(* IEC 61131-3 sources: Industry-PLC-LLM/data/PLCBEAD_repo/PLCBEAD_PLCEmbed-main/PLC-BEAD/Source/PLC_Programs (part 14) *)

(* ---- V3_XPRO.ST ---- *)
TYPE oscat_vector_3 :
	STRUCT
		X : REAL;
		Y : REAL;
		Z : REAL;
	END_STRUCT;
END_TYPE

FUNCTION_BLOCK V3_XPRO_Block
	VAR_INPUT
		A :	oscat_vector_3;
		B :	oscat_vector_3;
	END_VAR

	VAR_OUTPUT
		V3_XPRO :	oscat_vector_3;
	END_VAR

	V3_XPRO.X := A.Y * B.Z - A.Z * B.Y;
	V3_XPRO.Y := A.Z * B.X - A.X * B.Z;
	V3_XPRO.Z := A.X * B.Y - A.Y * B.X;

END_FUNCTION_BLOCK

PROGRAM program0
  	VAR
		A :	oscat_vector_3;
		B :	oscat_vector_3;
		V3_XPRO :	oscat_vector_3;
		func_block : V3_XPRO_Block;
  	END_VAR
	func_block.A := A;
	func_block.B := B;
	func_block();
	V3_XPRO := func_block.V3_XPRO;
END_PROGRAM

CONFIGURATION Config0
  RESOURCE Res0 ON PLC
    TASK task0(INTERVAL := T#20ms,PRIORITY := 0);
    PROGRAM instance0 WITH task0 : program0;
  END_RESOURCE
END_CONFIGURATION

(* ---- V3_YANG.ST ---- *)
TYPE oscat_vector_3:
  	STRUCT
		X : REAL;
		Y : REAL;
		Z : REAL;
  	END_STRUCT;
END_TYPE

FUNCTION_BLOCK V3_ABS_Block

	VAR_INPUT
		A :	oscat_vector_3;
	END_VAR

	VAR_OUTPUT
		V3_ABS :	REAL;
	END_VAR

	V3_ABS := SQRT(A.X * A.X + A.Y * A.Y + A.Z * A.Z);

END_FUNCTION_BLOCK

FUNCTION_BLOCK V3_YANG_Block
	VAR_INPUT
		A :	oscat_vector_3;
	END_VAR

	VAR_OUTPUT
		V3_YANG :	REAL;
	END_VAR

	VAR
		la :	REAL;
		V3_ABS :	V3_ABS_Block;
	END_VAR

	V3_ABS(A:=A);
	la:=V3_ABS.V3_ABS;

	IF la > 0.0 THEN
		V3_YANG := ACOS(A.Y / la);
	ELSE
		V3_YANG := 0.0;
	END_IF;

END_FUNCTION_BLOCK

PROGRAM program0
  	VAR
		A :	oscat_vector_3;
		V3_YANG :	REAL;
		func_block : V3_YANG_Block;
  	END_VAR
	func_block.A := A;
	func_block();
	V3_YANG := func_block.V3_YANG;
END_PROGRAM

CONFIGURATION Config0
  RESOURCE Res0 ON PLC
    TASK task0(INTERVAL := T#20ms,PRIORITY := 0);
    PROGRAM instance0 WITH task0 : program0;
  END_RESOURCE
END_CONFIGURATION

(* ---- V3_ZANG.ST ---- *)
TYPE oscat_vector_3:
  STRUCT
	X : REAL;
	Y : REAL;
	Z : REAL;
  END_STRUCT;
END_TYPE

FUNCTION_BLOCK V3_ABS_Block

	VAR_INPUT
		A :	oscat_vector_3;
	END_VAR

	VAR_OUTPUT
		V3_ABS :	REAL;
	END_VAR

	V3_ABS := SQRT(A.X * A.X + A.Y * A.Y + A.Z * A.Z);

END_FUNCTION_BLOCK

FUNCTION_BLOCK V3_ZANG_Block
	VAR_INPUT
		A :	oscat_vector_3;
	END_VAR

	VAR_OUTPUT
		V3_ZANG :	REAL;
	END_VAR

	VAR
		la :	REAL;
		V3_ABS :	V3_ABS_Block;
	END_VAR

	V3_ABS(A:=A);
	la:=V3_ABS.V3_ABS;

	IF la > 0.0 THEN
		V3_ZANG := ACOS(A.Z / la);
	ELSE
		V3_ZANG := 0.0;
	END_IF;

END_FUNCTION_BLOCK

PROGRAM program0
  	VAR
		A :	oscat_vector_3;
		V3_ZANG :	REAL;
		func_block : V3_ZANG_Block;
  	END_VAR
	func_block.A := A;
	func_block();
	V3_ZANG := func_block.V3_ZANG;
END_PROGRAM

CONFIGURATION Config0
  RESOURCE Res0 ON PLC
    TASK task0(INTERVAL := T#20ms,PRIORITY := 0);
    PROGRAM instance0 WITH task0 : program0;
  END_RESOURCE
END_CONFIGURATION

(* ---- WATER_CP.ST ---- *)
TYPE
	oscat_ARRAY_X               : ARRAY [0..1]    OF REAL;
	oscat_XY                    : ARRAY [1..20]   OF oscat_ARRAY_X := [0,0,0,0,0,0,0,0,0,0,0,0,0,0,0,0,0,0,0,0];
END_TYPE

FUNCTION_BLOCK LINEAR_INT_Block

	VAR_INPUT
		X :	REAL;
		XY :	oscat_XY;
		PTS :	INT;
	END_VAR

	VAR_OUTPUT
		LINEAR_INT :	REAL;
	END_VAR

	VAR
		i :	INT;
		i2 :	INT;
	END_VAR

	pts := MIN(pts,20);

	i := 2;

	WHILE (i < pts) AND (XY[i][0] < X) DO
		i := i + 1;
	END_WHILE;

	i2 := i-1;

	LINEAR_INT := ((XY[i][1] - XY[i2][1]) * X - XY[i][1] * XY[i2][0] + XY[i2][1] * XY[i][0]) / (XY[i][0] - XY[i2][0]);

END_FUNCTION_BLOCK

FUNCTION_BLOCK WATER_CP_Block

    VAR_INPUT
        T :	REAL;
    END_VAR

    VAR_OUTPUT
        CAP :	REAL;
    END_VAR

    VAR
        Pts :	INT;
        data :	oscat_XY;
        FB_LINEAR_INT :	LINEAR_INT_Block;
    END_VAR

    IF Pts = 0 THEN
        Pts := 10;

        data[01][0] := REAL#0.0;
        data[01][1] := REAL#4.228;
        data[02][0] := REAL#05.0;
        data[02][1] := REAL#4.200;
        data[03][0] := REAL#10.0;
        data[03][1] := REAL#4.188;
        data[04][0] := REAL#15.0;
        data[04][1] := REAL#4.184;
        data[05][0] := REAL#50.0;
        data[05][1] := REAL#4.181;
        data[06][0] := REAL#60.0;
        data[06][1] := REAL#4.183;
        data[07][0] := REAL#70.0;
        data[07][1] := REAL#4.187;
        data[08][0] := REAL#80.0;
        data[08][1] := REAL#4.194;
        data[09][0] := REAL#90.0;
        data[09][1] := REAL#4.204;
        data[10][0] := REAL#100.0;
        data[10][1] := REAL#4.220;

    END_IF;

    FB_LINEAR_INT(X:=T,XY:=Data,Pts:=Pts);
    cap:=FB_LINEAR_INT.LINEAR_INT;

END_FUNCTION_BLOCK

PROGRAM program0
	VAR
		T :	REAL;
        CAP :	REAL;

		func_block : WATER_CP_Block;
	END_VAR
	func_block.T := T;

	func_block();
	CAP  := func_block.CAP;
END_PROGRAM

CONFIGURATION Config0
	RESOURCE Res0 ON PLC
		TASK task0(INTERVAL := T#20ms,PRIORITY := 0);
		PROGRAM instance0 WITH task0 : program0;
	END_RESOURCE
END_CONFIGURATION

(* ---- WATER_ENTHALPY.ST ---- *)
TYPE
	oscat_ARRAY_X               : ARRAY [0..1]    OF REAL;
	oscat_XY                    : ARRAY [1..20]   OF oscat_ARRAY_X := [0,0,0,0,0,0,0,0,0,0,0,0,0,0,0,0,0,0,0,0];
END_TYPE

FUNCTION_BLOCK LINEAR_INT_Block

	VAR_INPUT
		X :	REAL;
		XY :	oscat_XY;
		PTS :	INT;
	END_VAR

	VAR_OUTPUT
		LINEAR_INT :	REAL;
	END_VAR

	VAR
		i :	INT;
		i2 :	INT;
	END_VAR

	pts := MIN(pts,20);

	i := 2;

	WHILE (i < pts) AND (XY[i][0] < X) DO
		i := i + 1;
	END_WHILE;

	i2 := i-1;

	LINEAR_INT := ((XY[i][1] - XY[i2][1]) * X - XY[i][1] * XY[i2][0] + XY[i2][1] * XY[i][0]) / (XY[i][0] - XY[i2][0]);

END_FUNCTION_BLOCK

FUNCTION_BLOCK WATER_ENTHALPY_Block

    VAR_INPUT
        T :	REAL;
    END_VAR

    VAR_OUTPUT
        RESULT :	REAL;
    END_VAR

    VAR
        Pts :	INT;
        data :	oscat_XY;
        FB_LINEAR_INT :	LINEAR_INT_Block;
    END_VAR

    IF Pts = 0 THEN
        Pts := 11;
        data[01][0] := REAL#0.0;
        data[01][1] := REAL#0.06;
        data[02][0] := REAL#10.0;
        data[02][1] := REAL#42.1;
        data[03][0] := REAL#20.0;
        data[03][1] := REAL#83.9;
        data[04][0] := REAL#30.0;
        data[04][1] := REAL#125.8;
        data[05][0] := REAL#40.0;
        data[05][1] := REAL#167.58;
        data[06][0] := REAL#50.0;
        data[06][1] := REAL#209.4;
        data[07][0] := REAL#60.0;
        data[07][1] := REAL#251.2;
        data[08][0] := REAL#70.0;
        data[08][1] := REAL#293.1;
        data[09][0] := REAL#80.0;
        data[09][1] := REAL#335.0;
        data[10][0] := REAL#90.0;
        data[10][1] := REAL#377.0;
        data[11][0] := REAL#100.0;
        data[11][1] := REAL#419.1;
    END_IF;

    FB_LINEAR_INT(X:=T,XY:=Data,Pts:=Pts);
    Result :=FB_LINEAR_INT.LINEAR_INT;

END_FUNCTION_BLOCK

PROGRAM program0
	VAR
		T :	REAL;
		RESULT :	REAL;

		func_block : WATER_ENTHALPY_Block;
	END_VAR
	func_block.T := T;

	func_block();
	RESULT  := func_block.RESULT;
END_PROGRAM

CONFIGURATION Config0
	RESOURCE Res0 ON PLC
		TASK task0(INTERVAL := T#20ms,PRIORITY := 0);
		PROGRAM instance0 WITH task0 : program0;
	END_RESOURCE
END_CONFIGURATION

(* ---- WEEKDAY_TO_STRING.ST ---- *)
TYPE
	oscat_STRING2 : STRING;
	oscat_STRING10 : STRING;
END_TYPE

TYPE oscat_HOLIDAY_DATA :
	STRUCT
		NAME : STRING;
		DAY : SINT;
		MONTH : SINT;
		USE : SINT;
		PAD_BYTE : BYTE;
	END_STRUCT;
END_TYPE

TYPE
	oscat_HOLIDAY_DATA_0_29 	: ARRAY [0..29] OF oscat_HOLIDAY_DATA;
END_TYPE

TYPE
	oscat_ELEMENT_WEEKDAYS	: ARRAY [1..7] OF oscat_STRING10;
  	oscat_WEEKDAYS			: ARRAY [1..3] OF oscat_ELEMENT_WEEKDAYS := [0,0,0];
	oscat_ELEMENT_WEEKDAYS2	: ARRAY [1..7] OF oscat_STRING2;
  	oscat_WEEKDAYS2			: ARRAY [1..3] OF oscat_ELEMENT_WEEKDAYS2 := [0,0,0];
END_TYPE

TYPE oscat_LANGUAGE:
  STRUCT
    DEFAULT 	: INT;
	LMAX    	: INT;
  END_STRUCT;
END_TYPE

FUNCTION_BLOCK SETUP_HOLIDAY_FR_Block

	VAR_IN_OUT
		HD :	oscat_HOLIDAY_DATA_0_29;
	END_VAR

	VAR
		init :	BOOL;
	END_VAR

	IF init THEN RETURN; END_IF;

	init := TRUE;

	HD[00].NAME := 'Nouve an';
	HD[00].DAY  := SINT#01;
	HD[00].MONTH := SINT#01;
	HD[00].USE := SINT#01;

	HD[01].NAME := 'St Valentin';
	HD[01].DAY  := SINT#14;
	HD[01].MONTH := SINT#02;
	HD[01].USE := SINT#00;

	HD[02].NAME := 'Vendredi Saint (alsace)';
	HD[02].DAY  := SINT#-2;
	HD[02].MONTH := SINT#00;
	HD[02].USE := SINT#00;

	HD[03].NAME := 'Dimanche de pques';
	HD[03].DAY  := SINT#00;
	HD[03].MONTH := SINT#00;
	HD[03].USE := SINT#01;

	HD[04].NAME := 'Lundi de pques';
	HD[04].DAY  := SINT#01;
	HD[04].MONTH := SINT#00;
	HD[04].USE := SINT#01;

	HD[05].NAME := 'Jeudi de Ascension';
	HD[05].DAY  := SINT#39;
	HD[05].MONTH := SINT#00;
	HD[05].USE := SINT#01;

	HD[06].NAME := 'dimanche de Pentecte';
	HD[06].DAY  := SINT#49;
	HD[06].MONTH := SINT#00;
	HD[06].USE := SINT#01;

	HD[07].NAME := 'jeudi de la Trinit';
	HD[07].DAY  := SINT#60;
	HD[07].MONTH := SINT#00;
	HD[07].USE := SINT#00;

	HD[08].NAME := 'Fte du travail';
	HD[08].DAY  := SINT#01;
	HD[08].MONTH := SINT#05;
	HD[08].USE := SINT#01;

	HD[09].NAME := 'Victoire 1945 ';
	HD[09].DAY  := SINT#08;
	HD[09].MONTH := SINT#05;
	HD[09].USE := SINT#01;

	HD[10].NAME := 'Prise de La bastille';
	HD[10].DAY  := SINT#14;
	HD[10].MONTH := SINT#07;
	HD[10].USE := SINT#01;

	HD[11].NAME := '15 Aot 1944';
	HD[11].DAY  := SINT#15;
	HD[11].MONTH := SINT#08;
	HD[11].USE := SINT#01;

	HD[12].NAME := 'Halloween';
	HD[12].DAY  := SINT#31;
	HD[12].MONTH := SINT#10;
	HD[12].USE := SINT#00;

	HD[13].NAME := 'Armistice 1918';
	HD[13].DAY  := SINT#11;
	HD[13].MONTH := SINT#11;
	HD[13].USE := SINT#01;

	HD[14].NAME := 'Nol';
	HD[14].DAY  := SINT#25;
	HD[14].MONTH := SINT#12;
	HD[14].USE := SINT#01;

	HD[15].NAME := 'Saint tienne (alsace)';
	HD[15].DAY  := SINT#26;
	HD[15].MONTH := SINT#12;
	HD[15].USE := SINT#00;

	HD[16].NAME := 'Fte de la musique';
	HD[16].DAY  := SINT#21;
	HD[16].MONTH := SINT#06;
	HD[16].USE := SINT#00;
END_FUNCTION_BLOCK

FUNCTION_BLOCK SETUP_LANGUAGE_Block

	VAR_IN_OUT
		LANGUAGE :	oscat_LANGUAGE;
	END_VAR

	VAR
		init :	BOOL;
	END_VAR

	IF init THEN RETURN; END_IF;
	init := TRUE;

	LANGUAGE.DEFAULT  := 1; (* 1=english, 2=german 3=french *)
	LANGUAGE.LMAX := 3;
END_FUNCTION_BLOCK

FUNCTION_BLOCK SETUP_WEEKDAYS_Block

	VAR_IN_OUT
		WEEKDAYS :	oscat_WEEKDAYS;
	END_VAR

	VAR
		init :	BOOL;
	END_VAR

	IF init THEN RETURN; END_IF;
	init := TRUE;

	WEEKDAYS[1][01] := 'Monday';
	WEEKDAYS[1][02] := 'Tuesday';
	WEEKDAYS[1][03] := 'Wednesday';
	WEEKDAYS[1][04] := 'Thursday';
	WEEKDAYS[1][05] := 'Friday';
	WEEKDAYS[1][06] := 'Saturday';
	WEEKDAYS[1][07] := 'Sunday';

	WEEKDAYS[2][01] := 'Montag';
	WEEKDAYS[2][02] := 'Dienstag';
	WEEKDAYS[2][03] := 'Mittwoch';
	WEEKDAYS[2][04] := 'Donnerstag';
	WEEKDAYS[2][05] := 'Freitag';
	WEEKDAYS[2][06] := 'Samstag';
	WEEKDAYS[2][07] := 'Sonntag';

	WEEKDAYS[3][01] := 'Lundi';
	WEEKDAYS[3][02] := 'Mardi';
	WEEKDAYS[3][03] := 'Mercredi';
	WEEKDAYS[3][04] := 'Jeudi';
	WEEKDAYS[3][05] := 'Vendredi';
	WEEKDAYS[3][06] := 'Samedi';
	WEEKDAYS[3][07] := 'Dimanche';
END_FUNCTION_BLOCK

FUNCTION_BLOCK WEEKDAY_TO_STRING_Block
	VAR_INPUT
		WDAY :	INT;
		LANG :	INT;
		LX :	INT;
	END_VAR

	VAR_OUTPUT
		WEEKDAY_TO_STRING :	STRING;
	END_VAR

	VAR
		LY :	INT;
		SETUP_LANGUAGE :	SETUP_LANGUAGE_Block;
		LANGUAGE :	oscat_LANGUAGE;
		WEEKDAYS :	oscat_WEEKDAYS;
		WEEKDAYS2 :	oscat_WEEKDAYS2;
		SETUP_WEEKDAYS :	SETUP_WEEKDAYS_Block;
		SETUP_WEEKDAYS2 :	SETUP_WEEKDAYS2_Block;
	END_VAR

	SETUP_WEEKDAYS(WEEKDAYS:=WEEKDAYS);
	WEEKDAYS:=SETUP_WEEKDAYS.WEEKDAYS;
	SETUP_WEEKDAYS2(WEEKDAYS2:=WEEKDAYS2);
	WEEKDAYS2:=SETUP_WEEKDAYS2.WEEKDAYS2;
	SETUP_LANGUAGE(LANGUAGE:=LANGUAGE);
	LANGUAGE:=SETUP_LANGUAGE.LANGUAGE;

	IF LANG = 0 THEN ly := LANGUAGE.DEFAULT; ELSE ly := MIN(LANG, LANGUAGE.LMAX); END_IF;
	IF wday < 1 OR wday > 7 THEN
		RETURN;
	ELSIF LX = 0 THEN
		WEEKDAY_TO_STRING := WEEKDAYS[ly][WDAY];
	ELSIF Lx = 2 THEN
		WEEKDAY_TO_STRING := WEEKDAYS2[ly][WDAY];
	END_IF;

END_FUNCTION_BLOCK

FUNCTION_BLOCK SETUP_WEEKDAYS2_Block

	VAR_IN_OUT
		WEEKDAYS2 :	oscat_WEEKDAYS2;
	END_VAR

	VAR
		init :	BOOL;
	END_VAR

	IF init THEN RETURN; END_IF;
	init := TRUE;

	WEEKDAYS2[1][01] := 'Mo';
	WEEKDAYS2[1][02] := 'Tu';
	WEEKDAYS2[1][03] := 'We';
	WEEKDAYS2[1][04] := 'Th';
	WEEKDAYS2[1][05] := 'Fr';
	WEEKDAYS2[1][06] := 'Sa';
	WEEKDAYS2[1][07] := 'Su';

	WEEKDAYS2[2][01] := 'Mo';
	WEEKDAYS2[2][02] := 'Di';
	WEEKDAYS2[2][03] := 'Mi';
	WEEKDAYS2[2][04] := 'Do';
	WEEKDAYS2[2][05] := 'Fr';
	WEEKDAYS2[2][06] := 'Sa';
	WEEKDAYS2[2][07] := 'So';

	WEEKDAYS2[3][01] := 'Lu';
	WEEKDAYS2[3][02] := 'Ma';
	WEEKDAYS2[3][03] := 'Me';
	WEEKDAYS2[3][04] := 'Je';
	WEEKDAYS2[3][05] := 'Ve';
	WEEKDAYS2[3][06] := 'Sa';
	WEEKDAYS2[3][07] := 'Di';
END_FUNCTION_BLOCK

PROGRAM program0
  	VAR
		WDAY :	INT;
		LANG :	INT;
		LX :	INT;
		WEEKDAY_TO_STRING :	STRING;
		func_block : WEEKDAY_TO_STRING_Block;
  	END_VAR
	func_block.WDAY := WDAY;
	func_block.LANG := LANG;
	func_block.LX := LX;
	func_block();
	WEEKDAY_TO_STRING := func_block.WEEKDAY_TO_STRING;
END_PROGRAM

CONFIGURATION Config0
  RESOURCE Res0 ON PLC
    TASK task0(INTERVAL := T#20ms,PRIORITY := 0);
    PROGRAM instance0 WITH task0 : program0;
  END_RESOURCE
END_CONFIGURATION

(* ---- ACOSH.ST ---- *)
FUNCTION ACOSH:REAL
	VAR_INPUT
		X :	REAL;
	END_VAR
	ACOSH := LN(SQRT(X * X - 1.0) + X);

END_FUNCTION

PROGRAM program0
  VAR
    LocalVar0 : REAL;
    LocalOUT  : REAL;
  END_VAR

  LocalOUT := ACOSH(LocalVar0);
END_PROGRAM

CONFIGURATION Config0
  RESOURCE Res0 ON PLC
    TASK task0(INTERVAL := T#20ms,PRIORITY := 0);
    PROGRAM instance0 WITH task0 : program0;
  END_RESOURCE
END_CONFIGURATION

(* ---- ACOTH.ST ---- *)
FUNCTION ACOTH:REAL
	VAR_INPUT
		X :	REAL;
	END_VAR

	ACOTH := LN((x+1.0)/(x-1.0))*0.5;

END_FUNCTION

PROGRAM program0
  VAR
    LocalVar0 : REAL;
    LocalOUT  : REAL;
  END_VAR

  LocalOUT := ACOTH(LocalVar0);
END_PROGRAM

CONFIGURATION Config0
  RESOURCE Res0 ON PLC
    TASK task0(INTERVAL := T#20ms,PRIORITY := 0);
    PROGRAM instance0 WITH task0 : program0;
  END_RESOURCE
END_CONFIGURATION

(* ---- AGDF.ST ---- *)
FUNCTION AGDF:REAL
	VAR_INPUT
		X :	REAL;
	END_VAR

	AGDF := LN((1.0 + SIN(X)) / COS(X));
END_FUNCTION

PROGRAM program0
  VAR
    LocalVar0 : REAL;
    LocalOUT  : REAL;
  END_VAR

  LocalOUT := AGDF(LocalVar0);
END_PROGRAM

CONFIGURATION Config0
  RESOURCE Res0 ON PLC
    TASK task0(INTERVAL := T#20ms,PRIORITY := 0);
    PROGRAM instance0 WITH task0 : program0;
  END_RESOURCE
END_CONFIGURATION

(* ---- AIN.ST ---- *)
FUNCTION _BYTE_TO_INT:INT
	VAR_INPUT
		IN :	BYTE;
	END_VAR

	_BYTE_TO_INT := USINT_TO_INT(BYTE_TO_USINT(IN));
END_FUNCTION

FUNCTION _DWORD_TO_REAL:REAL
	VAR_INPUT
		IN :	DWORD;
	END_VAR

	_DWORD_TO_REAL := UDINT_TO_REAL(DWORD_TO_UDINT(IN));
END_FUNCTION

FUNCTION BIT_OF_DWORD:BOOL
	VAR_INPUT
		IN :	DWORD;
		N :	INT;
	END_VAR
	BIT_OF_DWORD := (SHR(in,n) AND DWORD#1) > DWORD#0;
END_FUNCTION

FUNCTION AIN:REAL
	VAR_INPUT
		IN :	DWORD;
		BITS :	BYTE;
		SIGN :	BYTE;
		LOW :	REAL;
		HIGH :	REAL;
	END_VAR

	VAR
		temp1 :	DWORD;
		temp2 :	DWORD;
		sx :	BOOL;
	END_VAR

	IF sign < BYTE#32 THEN
		temp1 := SHR(in, _BYTE_TO_INT(sign));
		sx := BIT_OF_DWORD(temp1,0); (* temp1.X0 *)
	ELSE
		sx := FALSE;
	END_IF;
	temp1 := SHR(DWORD#16#FFFFFFFF,32 - _BYTE_TO_INT(bits));
	temp2 := in AND temp1;
	AIN := (high - low)* _DWORD_TO_REAL(temp2) / _DWORD_TO_REAL(temp1) + low;
	IF sx THEN AIN := -AIN; END_IF;
END_FUNCTION

PROGRAM program0
  VAR
    LocalVar0 : DWORD;
	LocalVar1 : BYTE;
	LocalVar2 : BYTE;
	LocalVar3 : REAL;
	LocalVar4 : REAL;
    LocalOUT  : REAL;
  END_VAR

  LocalOUT := AIN(LocalVar0, LocalVar1, LocalVar2, LocalVar3, LocalVar4);
END_PROGRAM

CONFIGURATION Config0
  RESOURCE Res0 ON PLC
    TASK task0(INTERVAL := T#20ms,PRIORITY := 0);
    PROGRAM instance0 WITH task0 : program0;
  END_RESOURCE
END_CONFIGURATION

(* ---- AIR_DENSITY.ST ---- *)
FUNCTION SDD:REAL

	VAR_INPUT
		T :	REAL;
		ICE :	BOOL;
	END_VAR

	IF ice THEN
		SDD := 611.153 * EXP(22.4433 * T / (272.186 + T));
	ELSE
		SDD := 611.213 * EXP(17.5043 * T / (241.2 + T));
	END_IF;

END_FUNCTION

FUNCTION AIR_DENSITY:REAL

	VAR_INPUT
		T :	REAL;
		P :	REAL;
		RH :	REAL;
	END_VAR

	AIR_DENSITY := 101325.0 * (1.0 - RH * SDD(T, TRUE) * 3.773319E-3 / P) / (287.05 * ( T - -273.15));

END_FUNCTION

PROGRAM program0
  VAR
    T :	REAL;
	P :	REAL;
	RH :	REAL;
    CEIL5_OUT : REAL;
  END_VAR

  CEIL5_OUT := AIR_DENSITY(T, P, RH);
END_PROGRAM

CONFIGURATION Config0

  RESOURCE Res0 ON PLC
    TASK task0(INTERVAL := T#20ms,PRIORITY := 0);
    PROGRAM instance0 WITH task0 : program0;
  END_RESOURCE
END_CONFIGURATION

(* ---- AIR_ENTHALPY.ST ---- *)
FUNCTION SDD:REAL

	VAR_INPUT
		T :	REAL;
		ICE :	BOOL;
	END_VAR

	IF ice THEN
		SDD := 611.153 * EXP(22.4433 * T / (272.186 + T));
	ELSE
		SDD := 611.213 * EXP(17.5043 * T / (241.2 + T));
	END_IF;

END_FUNCTION

FUNCTION DEW_CON:REAL

	VAR_INPUT
		RH :	REAL;
		T :	REAL;
	END_VAR

	IF RH > 0.0 AND T > -50.0 THEN
		DEW_CON := 2.166824303E-2 * RH * SDD(T,FALSE)  / (T - -273.15);
	ELSE
		DEW_CON := 0.0;
	END_IF;

END_FUNCTION

FUNCTION AIR_ENTHALPY:REAL

	VAR_INPUT
		T :	REAL;
		RH :	REAL;
	END_VAR

	Air_enthalpy := 1.00482 * T + (1.86 * T + 2500.78) * dew_con(RH,T);

END_FUNCTION

PROGRAM program0
  VAR
    T :	REAL;
	RH :	REAL;
    CEIL5_OUT : REAL;
  END_VAR

  CEIL5_OUT := AIR_ENTHALPY(T, RH);
END_PROGRAM

CONFIGURATION Config0

  RESOURCE Res0 ON PLC
    TASK task0(INTERVAL := T#20ms,PRIORITY := 0);
    PROGRAM instance0 WITH task0 : program0;
  END_RESOURCE
END_CONFIGURATION

(* ---- AOUT.ST ---- *)
FUNCTION _DWORD_TO_REAL:REAL
	VAR_INPUT
		IN :	DWORD;
	END_VAR

	_DWORD_TO_REAL := UDINT_TO_REAL(DWORD_TO_UDINT(IN));
END_FUNCTION

FUNCTION SIGN_R : BOOL
  VAR_INPUT
    IN : REAL;
  END_VAR
  SIGN_R := in < 0.0;
END_FUNCTION

FUNCTION _REAL_TO_DWORD: DWORD

  VAR_INPUT
    X :	REAL;
  END_VAR

  IF REAL_TO_DWORD(0.5) = DWORD#1 THEN
    _REAL_TO_DWORD := REAL_TO_DWORD(x);
  ELSIF X > 0.0 THEN
    _REAL_TO_DWORD := REAL_TO_DWORD(x+0.5);
  ELSIF X < 0.0 THEN
    _REAL_TO_DWORD := REAL_TO_DWORD(x-0.5);
  ELSE
    _REAL_TO_DWORD := DWORD#0;
  END_IF;
END_FUNCTION

FUNCTION _BYTE_TO_INT:INT
	VAR_INPUT
		IN :	BYTE;
	END_VAR

	_BYTE_TO_INT := USINT_TO_INT(BYTE_TO_USINT(IN));
END_FUNCTION

FUNCTION AOUT:DWORD
	VAR_INPUT
		IN :	REAL;
		BITS :	BYTE;
		SIGN :	BYTE;
		LOW :	REAL;
		HIGH :	REAL;
	END_VAR

	VAR
		in2 :	REAL;
		sx :	BOOL;
	END_VAR

	IF sign < BYTE#32 THEN
		sx := sign_R(in);
		in2 := ABS(in);
	ELSE
		in2 := in;
	END_IF;

	in2 := LIMIT(low, in2, high);

	Aout := _REAL_TO_DWORD((in2 - low) / (high - low) * (_DWORD_TO_REAL(SHL(DWORD#2#1,_BYTE_TO_INT(bits))) - 1.0)   );
	IF sx THEN Aout := SHL(DWORD#2#1,_BYTE_TO_INT(sign)) OR Aout; END_IF;

END_FUNCTION

PROGRAM program0
  VAR
    LocalVar0 : REAL;
	LocalVar1 : BYTE;
	LocalVar2 : BYTE;
	LocalVar3 : REAL;
	LocalVar4 : REAL;
	LocalOUT  : DWORD;
  END_VAR
  	LocalOUT := AOUT(LocalVar0, LocalVar1, LocalVar2, LocalVar3,LocalVar4);
END_PROGRAM

CONFIGURATION Config0
  RESOURCE Res0 ON PLC
    TASK task0(INTERVAL := T#20ms,PRIORITY := 0);
    PROGRAM instance0 WITH task0 : program0;
  END_RESOURCE
END_CONFIGURATION

(* ---- AOUT1.ST ---- *)
FUNCTION SIGN_R : BOOL
  VAR_INPUT
    IN : REAL;
  END_VAR

  SIGN_R := in < 0.0;
END_FUNCTION

FUNCTION _REAL_TO_DWORD: DWORD

  VAR_INPUT
    X :	REAL;
  END_VAR

  IF REAL_TO_DWORD(0.5) = DWORD#1 THEN
    _REAL_TO_DWORD := REAL_TO_DWORD(x);
  ELSIF X > 0.0 THEN
    _REAL_TO_DWORD := REAL_TO_DWORD(x+0.5);
  ELSIF X < 0.0 THEN
    _REAL_TO_DWORD := REAL_TO_DWORD(x-0.5);
  ELSE
    _REAL_TO_DWORD := DWORD#0;
  END_IF;
END_FUNCTION

FUNCTION AOUT1:DWORD

	VAR_INPUT
		IN :	REAL;
		BIT_0 :	INT;
		BIT_N :	INT;
		SIGN :	INT;
		LOW :	REAL;
		HIGH :	REAL;
	END_VAR

	VAR
		in2 :	REAL;
		sx :	BOOL;
	END_VAR

	IF sign < 32 THEN
		sx := sign_R(in);
		in2 := ABS(in);
	ELSE
		sx := FALSE;
		in2 := in;
	END_IF;

	in2 := LIMIT_REAL(low, in2, high);

	AOUT1 :=  SHL(_REAL_TO_DWORD((in2 - low) / (high - low) * UDINT_TO_REAL(DWORD_TO_UDINT(SHL(DWORD#2#1,bit_n - Bit_0 + 1)) - UDINT#1)),Bit_0);

	IF sx THEN AOUT1 := SHL(DWORD#2#1,sign) OR AOUT1; END_IF;

END_FUNCTION

PROGRAM program0
  VAR
    LocalVar0 : REAL;
	LocalVar1 : INT;
	LocalVar21 : INT;
	LocalVar2 : INT;
	LocalVar3 : REAL;
	LocalVar4 : REAL;
	LocalOUT  : DWORD;
  END_VAR
  	LocalOUT := AOUT1(LocalVar0, LocalVar1,LocalVar21, LocalVar2, LocalVar3,LocalVar4);
END_PROGRAM

CONFIGURATION Config0
  RESOURCE Res0 ON PLC
    TASK task0(INTERVAL := T#20ms,PRIORITY := 0);
    PROGRAM instance0 WITH task0 : program0;
  END_RESOURCE
END_CONFIGURATION

(* ---- ASINH.ST ---- *)
FUNCTION ASINH:REAL
	VAR_INPUT
		X :	REAL;
	END_VAR

	ASINH := LN(SQRT(X * X + 1.0)+X);
END_FUNCTION

PROGRAM program0
  VAR
    LocalVar0 : REAL;
    LocalOUT  : REAL;
  END_VAR

  LocalOUT := ASINH(LocalVar0);
END_PROGRAM

CONFIGURATION Config0
  RESOURCE Res0 ON PLC
    TASK task0(INTERVAL := T#20ms,PRIORITY := 0);
    PROGRAM instance0 WITH task0 : program0;
  END_RESOURCE
END_CONFIGURATION

(* ---- ATAN2.ST ---- *)
FUNCTION ATAN2:REAL
	VAR_INPUT
		X :	REAL;
		Y :	REAL;
	END_VAR

	IF X > 0.0 THEN
		ATAN2 := ATAN(Y/X);
	ELSIF X < 0.0 THEN
		IF Y >= 0.0 THEN
			ATAN2 := ATAN(Y/X) + 3.14159265358979323846264338327950288;
		ELSE
			ATAN2 := ATAN(Y/X) - 3.14159265358979323846264338327950288;
		END_IF;
	ELSIF Y > 0.0 THEN
		ATAN2 := 1.5707963267948965580;
	ELSIF Y < 0.0 THEN
		ATAN2 := -1.5707963267948965580;
	ELSE
		ATAN2 := 0.0;
	END_IF;

END_FUNCTION

PROGRAM program0
  VAR
    LocalVar0 : REAL;
	LocalVar1 : REAL;
    LocalOUT  : REAL;
  END_VAR

  LocalOUT := ATAN2(LocalVar0, LocalVar1);
END_PROGRAM

CONFIGURATION Config0
  RESOURCE Res0 ON PLC
    TASK task0(INTERVAL := T#20ms,PRIORITY := 0);
    PROGRAM instance0 WITH task0 : program0;
  END_RESOURCE
END_CONFIGURATION

(* ---- ATANH.ST ---- *)
FUNCTION ATANH:REAL
	VAR_INPUT
		X :	REAL;
	END_VAR

	ATANH := LN((1.0 + x)/(1.0 - x)) * 0.5;

END_FUNCTION

PROGRAM program0
  VAR
    LocalVar0 : REAL;
    LocalOUT  : REAL;
  END_VAR

  LocalOUT := ATANH(LocalVar0);
END_PROGRAM

CONFIGURATION Config0
  RESOURCE Res0 ON PLC
    TASK task0(INTERVAL := T#20ms,PRIORITY := 0);
    PROGRAM instance0 WITH task0 : program0;
  END_RESOURCE
END_CONFIGURATION

(* ---- BAND_B.ST ---- *)
FUNCTION BAND_B:BYTE
	VAR_INPUT
		X :	BYTE;
		B :	BYTE;
	END_VAR

	IF X < B THEN
		BAND_B := BYTE#0;
	ELSIF X > USINT_TO_BYTE(USINT#255 - BYTE_TO_USINT(B)) THEN
		BAND_B := BYTE#255;
	ELSE
		BAND_B := X;
	END_IF;
END_FUNCTION
PROGRAM program0
  VAR
    LocalVar0 : BYTE;
	LocalVar1 : BYTE;
    LocalOUT  : BYTE;
  END_VAR

  LocalOUT := BAND_B(LocalVar0, LocalVar1);
END_PROGRAM

CONFIGURATION Config0
  RESOURCE Res0 ON PLC
    TASK task0(INTERVAL := T#20ms,PRIORITY := 0);
    PROGRAM instance0 WITH task0 : program0;
  END_RESOURCE
END_CONFIGURATION

(* ---- BCDC_TO_INT.ST ---- *)
FUNCTION _BYTE_TO_INT:INT
	VAR_INPUT
		IN :	BYTE;
	END_VAR

	_BYTE_TO_INT := USINT_TO_INT(BYTE_TO_USINT(IN));

END_FUNCTION

FUNCTION BCDC_TO_INT:INT
	VAR_INPUT
		IN :	BYTE;
	END_VAR

	BCDC_TO_INT := _BYTE_TO_INT(in AND BYTE#16#0F) + (_BYTE_TO_INT(SHR(in,4)) * 10);
END_FUNCTION

PROGRAM program0
  VAR
    LocalVar0 : BYTE;
    LocalOUT  : INT;
  END_VAR

  LocalOUT := BCDC_TO_INT(LocalVar0);
END_PROGRAM

CONFIGURATION Config0
  RESOURCE Res0 ON PLC
    TASK task0(INTERVAL := T#20ms,PRIORITY := 0);
    PROGRAM instance0 WITH task0 : program0;
  END_RESOURCE
END_CONFIGURATION

(* ---- BETA.ST ---- *)
FUNCTION GAMMA:REAL
	VAR_INPUT
		X :	REAL;
	END_VAR

	IF x > 0.0 THEN
		GAMMA := SQRT(6.28318530717958647692528676655900576 / X) * EXPT(0.367879441171442 * (x + 1.0 / (12.0 * x - 0.1 / X)), X);
	END_IF;
END_FUNCTION

FUNCTION BETA:REAL

	VAR_INPUT
		X :	REAL;
		Y :	REAL;
	END_VAR

	BETA := GAMMA(X)*GAMMA(Y) / GAMMA(x+y);

END_FUNCTION

PROGRAM program0
  VAR
    LocalVar0 : REAL;
	LocalVar1 : REAL;
    LocalOUT  : REAL;
  END_VAR

  LocalOUT := BETA(LocalVar0, LocalVar1);
END_PROGRAM

CONFIGURATION Config0
  RESOURCE Res0 ON PLC
    TASK task0(INTERVAL := T#20ms,PRIORITY := 0);
    PROGRAM instance0 WITH task0 : program0;
  END_RESOURCE
END_CONFIGURATION

(* ---- BFT_TO_MS.ST ---- *)
FUNCTION BFT_TO_MS:REAL
	VAR_INPUT
		BFT :	INT;
	END_VAR

	BFT_TO_MS := EXPT(INT_TO_REAL(BFT), 1.5) * 0.836;

END_FUNCTION

PROGRAM program0
  VAR
    LocalVar0 : INT;
    LocalOUT  : REAL;
  END_VAR

  LocalOUT := BFT_TO_MS(LocalVar0);
END_PROGRAM

CONFIGURATION Config0
  RESOURCE Res0 ON PLC
    TASK task0(INTERVAL := T#20ms,PRIORITY := 0);
    PROGRAM instance0 WITH task0 : program0;
  END_RESOURCE
END_CONFIGURATION

(* ---- BINOM.ST ---- *)
FUNCTION BINOM:INT
	VAR_INPUT
		N :	INT;
		K :	INT;
	END_VAR

	VAR
		i :	INT;
		N2 :	INT;
		K2 :	INT;
	END_VAR

	K2 := K;
	N2 := N;
	IF 2 * K2 > N2 THEN
		K2 := N2 - K2;
	END_IF;
	IF K2 > N2 THEN
		RETURN;
	ELSIF K2 = 0 OR K2 = N2 THEN
		BINOM := 1;
	ELSIF K2 = 1 THEN
		BINOM := N2;
	ELSE
		BINOM := N2;
		N2 := N2 + 1;
		FOR i := 2 TO K2 DO
			BINOM := BINOM * (N2 - i) / i;
		END_FOR;
	END_IF;
END_FUNCTION

PROGRAM program0
  VAR
    LocalVar0 : INT;
	LocalVar1 : INT;
    LocalOUT  : INT;
  END_VAR

  LocalOUT := BINOM(LocalVar0, LocalVar1);
END_PROGRAM

CONFIGURATION Config0
  RESOURCE Res0 ON PLC
    TASK task0(INTERVAL := T#20ms,PRIORITY := 0);
    PROGRAM instance0 WITH task0 : program0;
  END_RESOURCE
END_CONFIGURATION

(* ---- BIT_COUNT.ST ---- *)
FUNCTION BIT_COUNT:INT

	VAR_INPUT
		IN :	DWORD;
	END_VAR

	VAR
		in_temp :	DWORD;
	END_VAR

	in_temp := IN;
	WHILE in_temp > DWORD#0 DO
		IF (in_temp AND DWORD#16#00000001) > DWORD#0 THEN Bit_Count := Bit_Count +1; END_IF;
		in_temp := SHR(in_temp,1);
	END_WHILE;

END_FUNCTION

PROGRAM program0
  VAR
    LocalVar0 : DWORD;
    LocalOUT  : INT;
  END_VAR

  LocalOUT := BIT_COUNT(LocalVar0);
END_PROGRAM

CONFIGURATION Config0
  RESOURCE Res0 ON PLC
    TASK task0(INTERVAL := T#20ms,PRIORITY := 0);
    PROGRAM instance0 WITH task0 : program0;
  END_RESOURCE
END_CONFIGURATION

(* ---- BIT_LOAD_B.ST ---- *)
FUNCTION BIT_LOAD_B:BYTE
	VAR_INPUT
		IN :	BYTE;
		VAL :	BOOL;
		POS :	INT;
	END_VAR

	IF VAL THEN
		BIT_LOAD_B := in OR SHL(BYTE#1,pos);
	ELSE
		BIT_LOAD_B := in AND (NOT SHL(BYTE#1,pos));
	END_IF;
END_FUNCTION

PROGRAM program0
  VAR
    LocalVar0 : BYTE;
	LocalVar1 : BOOL;
	LocalVar2 : INT;
    LocalOUT  : BYTE;
  END_VAR

  LocalOUT := BIT_LOAD_B(LocalVar0, LocalVar1, LocalVar2);
END_PROGRAM

CONFIGURATION Config0
  RESOURCE Res0 ON PLC
    TASK task0(INTERVAL := T#20ms,PRIORITY := 0);
    PROGRAM instance0 WITH task0 : program0;
  END_RESOURCE
END_CONFIGURATION

(* ---- BIT_LOAD_B2.ST ---- *)
FUNCTION BIT_LOAD_B2:BYTE
	VAR_INPUT
		I :	BYTE;
		D :	BOOL;
		P :	INT;
		N :	INT;
	END_VAR

	IF D THEN
		BIT_LOAD_B2 := ROL(SHR(BYTE#255, 8 - N) OR ROR(I, P), P);
	ELSE
		BIT_LOAD_B2 := ROL(SHL(BYTE#255, N) AND ROR(I, P), P);
	END_IF;
END_FUNCTION

PROGRAM program0
  VAR
    LocalVar0 : BYTE;
	LocalVar1 : BOOL;
	LocalVar2 : INT;
	LocalVar3 : INT;
    LocalOUT  : BYTE;
  END_VAR

  LocalOUT := BIT_LOAD_B2(LocalVar0, LocalVar1, LocalVar2, LocalVar3);
END_PROGRAM

CONFIGURATION Config0
  RESOURCE Res0 ON PLC
    TASK task0(INTERVAL := T#20ms,PRIORITY := 0);
    PROGRAM instance0 WITH task0 : program0;
  END_RESOURCE
END_CONFIGURATION

(* ---- BIT_LOAD_DW.ST ---- *)
FUNCTION BIT_LOAD_DW:DWORD

	VAR_INPUT
		IN :	DWORD;
		VAL :	BOOL;
		POS :	INT;
	END_VAR

	IF val THEN
		BIT_LOAD_DW := in OR SHL(DWORD#1,pos);
	ELSE
		BIT_LOAD_DW := in AND (NOT SHL(DWORD#1,pos));
	END_IF;

END_FUNCTION

PROGRAM program0
  VAR
    LocalVar0 : DWORD;
	LocalVar1 : BOOL;
	LocalVar2 : INT;
    LocalOUT  : DWORD;
  END_VAR

  LocalOUT := BIT_LOAD_DW(LocalVar0, LocalVar1, LocalVar2);
END_PROGRAM

CONFIGURATION Config0
  RESOURCE Res0 ON PLC
    TASK task0(INTERVAL := T#20ms,PRIORITY := 0);
    PROGRAM instance0 WITH task0 : program0;
  END_RESOURCE
END_CONFIGURATION

(* ---- BIT_LOAD_DW2.ST ---- *)
FUNCTION BIT_LOAD_DW2:DWORD
	VAR_INPUT
		I :	DWORD;
		D :	BOOL;
		P :	INT;
		N :	INT;
	END_VAR

	IF D THEN
		BIT_LOAD_DW2 := ROL(SHR(DWORD#16#FFFFFFFF, 32 - N) OR ROR(I, P), P);
	ELSE
		BIT_LOAD_DW2 := ROL(SHL(DWORD#16#FFFFFFFF, N) AND ROR(I, P), P);
	END_IF;

END_FUNCTION

PROGRAM program0
  VAR
    LocalVar0 : DWORD;
	LocalVar1 : BOOL;
	LocalVar2 : INT;
	LocalVar3 : INT;
    LocalOUT  : DWORD;
  END_VAR

  LocalOUT := BIT_LOAD_DW2(LocalVar0, LocalVar1, LocalVar2, LocalVar3);
END_PROGRAM

CONFIGURATION Config0
  RESOURCE Res0 ON PLC
    TASK task0(INTERVAL := T#20ms,PRIORITY := 0);
    PROGRAM instance0 WITH task0 : program0;
  END_RESOURCE
END_CONFIGURATION

(* ---- BIT_LOAD_W.ST ---- *)
FUNCTION BIT_LOAD_W:WORD
	VAR_INPUT
		IN :	WORD;
		VAL :	BOOL;
		POS :	INT;
	END_VAR

	IF VAL THEN
		BIT_LOAD_W := in OR SHL(WORD#1,pos);
	ELSE
		BIT_LOAD_W := in AND (NOT SHL(WORD#1,pos));
	END_IF;
END_FUNCTION

PROGRAM program0
  VAR
    LocalVar0 : WORD;
	LocalVar1 : BOOL;
	LocalVar2 : INT;
    LocalOUT  : WORD;
  END_VAR

  LocalOUT := BIT_LOAD_W(LocalVar0, LocalVar1, LocalVar2);
END_PROGRAM

CONFIGURATION Config0
  RESOURCE Res0 ON PLC
    TASK task0(INTERVAL := T#20ms,PRIORITY := 0);
    PROGRAM instance0 WITH task0 : program0;
  END_RESOURCE
END_CONFIGURATION

(* ---- BIT_LOAD_W2.ST ---- *)
FUNCTION BIT_LOAD_W2:WORD
	VAR_INPUT
		I :	WORD;
		D :	BOOL;
		P :	INT;
		N :	INT;
	END_VAR

	IF D THEN
		BIT_LOAD_W2 := ROL(SHR(WORD#16#FFFF, 16 - N) OR ROR(I, P), P);
	ELSE
		BIT_LOAD_W2 := ROL(SHL(WORD#16#FFFF, N) AND ROR(I, P), P);
	END_IF;
END_FUNCTION

PROGRAM program0
  VAR
    LocalVar0 : WORD;
	LocalVar1 : BOOL;
	LocalVar2 : INT;
	LocalVar3 : INT;
    LocalOUT  : WORD;
  END_VAR

  LocalOUT := BIT_LOAD_W2(LocalVar0, LocalVar1, LocalVar2, LocalVar3);
END_PROGRAM

CONFIGURATION Config0
  RESOURCE Res0 ON PLC
    TASK task0(INTERVAL := T#20ms,PRIORITY := 0);
    PROGRAM instance0 WITH task0 : program0;
  END_RESOURCE
END_CONFIGURATION

(* ---- BIT_OF_DWORD.ST ---- *)
FUNCTION BIT_OF_DWORD : BOOL
  VAR_INPUT
    IN : DWORD;
    N : INT;
  END_VAR

  BIT_OF_DWORD := (SHR(in,N) AND 16#00000001) > 0;
END_FUNCTION

PROGRAM program0
  VAR
    LocalVar0 : DWORD;
    LocalVar2 : INT;
    LocalVar1 : BOOL;
    CEIL5_OUT : BOOL;
  END_VAR

  CEIL5_OUT := BIT_OF_DWORD(LocalVar0, LocalVar2);
  LocalVar1 := CEIL5_OUT;
END_PROGRAM

CONFIGURATION Config0

  RESOURCE Res0 ON PLC
    TASK task0(INTERVAL := T#20ms,PRIORITY := 0);
    PROGRAM instance0 WITH task0 : program0;
  END_RESOURCE
END_CONFIGURATION

(* ---- BIT_TOGGLE_B.ST ---- *)
FUNCTION BIT_TOGGLE_B:BYTE
	VAR_INPUT
		IN :	BYTE;
		POS :	INT;
	END_VAR

	BIT_TOGGLE_B := SHL(BYTE#1, POS) XOR IN;
END_FUNCTION

PROGRAM program0
  VAR
    LocalVar0 : BYTE;
    LocalVar1 : INT;
    CEIL5_OUT : BYTE;
  END_VAR

  CEIL5_OUT := BIT_TOGGLE_B(LocalVar0, LocalVar1);
END_PROGRAM

CONFIGURATION Config0

  RESOURCE Res0 ON PLC
    TASK task0(INTERVAL := T#20ms,PRIORITY := 0);
    PROGRAM instance0 WITH task0 : program0;
  END_RESOURCE
END_CONFIGURATION

(* ---- BIT_TOGGLE_DW.ST ---- *)
FUNCTION BIT_TOGGLE_DW:DWORD
	VAR_INPUT
		IN :	DWORD;
		POS :	INT;
	END_VAR

	BIT_TOGGLE_DW := SHL(DWORD#1, POS) XOR IN;

END_FUNCTION

PROGRAM program0
  VAR
    LocalVar0 : DWORD;
    LocalVar1 : INT;
    CEIL5_OUT : DWORD;
  END_VAR

  CEIL5_OUT := BIT_TOGGLE_DW(LocalVar0, LocalVar1);
END_PROGRAM

CONFIGURATION Config0

  RESOURCE Res0 ON PLC
    TASK task0(INTERVAL := T#20ms,PRIORITY := 0);
    PROGRAM instance0 WITH task0 : program0;
  END_RESOURCE
END_CONFIGURATION

(* ---- BIT_TOGGLE_W.ST ---- *)
FUNCTION BIT_TOGGLE_W:WORD
	VAR_INPUT
		IN :	WORD;
		POS :	INT;
	END_VAR

	BIT_TOGGLE_W := SHL(WORD#1, POS) XOR IN;
END_FUNCTION

PROGRAM program0
  VAR
    LocalVar0 : WORD;
    LocalVar1 : INT;
    CEIL5_OUT : WORD;
  END_VAR

  CEIL5_OUT := BIT_TOGGLE_W(LocalVar0, LocalVar1);
END_PROGRAM

CONFIGURATION Config0

  RESOURCE Res0 ON PLC
    TASK task0(INTERVAL := T#20ms,PRIORITY := 0);
    PROGRAM instance0 WITH task0 : program0;
  END_RESOURCE
END_CONFIGURATION

(* ---- BUILDING_VERSION.ST ---- *)
FUNCTION _INT_TO_UDINT:UDINT
	VAR_INPUT
		IN :	INT;
	END_VAR

	_INT_TO_UDINT := DINT_TO_UDINT(INT_TO_DINT(IN));
END_FUNCTION

FUNCTION SET_DATE:UDINT

	VAR_INPUT
		YEAR :	INT;
		MONTH :	INT;
		DAY :	INT;
	END_VAR

	VAR
		count :	INT;
	END_VAR

	IF month > 2 THEN
		count := (month - 1) * 30;
		IF month > 7 THEN
			count := count + DWORD_TO_INT(SHR(DINT_TO_DWORD(INT_TO_DINT(month) - INT_TO_DINT(3)),1));
		ELSE
			count := count + DWORD_TO_INT(SHR(DINT_TO_DWORD(INT_TO_DINT(month) - INT_TO_DINT(4)),1));
		END_IF;
		IF SHL(INT_TO_WORD(year),14) = WORD#0 THEN
			count := count + 1;
		END_IF;
	ELSE
		count := (month - 1) * 31;
	END_IF;
	SET_DATE := (_INT_TO_UDINT(count + day - 1) + DWORD_TO_UDINT(SHR(UDINT_TO_DWORD(_INT_TO_UDINT(year) * UDINT#1461 - UDINT#2878169), 2))) * UDINT#86400;

END_FUNCTION

FUNCTION BUILDING_VERSION:DWORD

	VAR_INPUT
		IN :	BOOL;
	END_VAR

	IF in THEN
		BUILDING_VERSION := UDINT_TO_DWORD(set_Date(2011,02,03));
	ELSE
		BUILDING_VERSION := DWORD#100;
	END_IF;

END_FUNCTION

PROGRAM program0
	VAR
		IN :	BOOL;
		CEIL5_OUT : DWORD;
	END_VAR

  	CEIL5_OUT := BUILDING_VERSION(IN);
END_PROGRAM

CONFIGURATION Config0

  RESOURCE Res0 ON PLC
    TASK task0(INTERVAL := T#20ms,PRIORITY := 0);
    PROGRAM instance0 WITH task0 : program0;
  END_RESOURCE
END_CONFIGURATION

(* ---- BYTE_OF_BIT.ST ---- *)
FUNCTION BYTE_OF_BIT:BYTE
	VAR_INPUT
		B0 :	BOOL;
		B1 :	BOOL;
		B2 :	BOOL;
		B3 :	BOOL;
		B4 :	BOOL;
		B5 :	BOOL;
		B6 :	BOOL;
		B7 :	BOOL;
	END_VAR
	Byte_of_bit := SHL(SHL(SHL(SHL(SHL(SHL(SHL(BOOL_TO_BYTE(B7),1) OR BOOL_TO_BYTE(B6),1)
	OR BOOL_TO_BYTE(B5),1) OR BOOL_TO_BYTE(B4),1) OR BOOL_TO_BYTE(B3),1) OR BOOL_TO_BYTE(B2),1)
	OR BOOL_TO_BYTE(B1),1) OR BOOL_TO_BYTE(B0);
END_FUNCTION

PROGRAM program0
  VAR
	B0 :	BOOL;
	B1 :	BOOL;
	B2 :	BOOL;
	B3 :	BOOL;
	B4 :	BOOL;
	B5 :	BOOL;
	B6 :	BOOL;
	B7 :	BOOL;
    LocalOUT  : BYTE;
  END_VAR

  LocalOUT := BYTE_OF_BIT(B0, B1, B2, B3, B4, B5, B6, B7);
END_PROGRAM

CONFIGURATION Config0
  RESOURCE Res0 ON PLC
    TASK task0(INTERVAL := T#20ms,PRIORITY := 0);
    PROGRAM instance0 WITH task0 : program0;
  END_RESOURCE
END_CONFIGURATION

(* ---- BYTE_OF_DWORD.ST ---- *)
FUNCTION _BYTE_TO_INT:INT
	VAR_INPUT
		IN :	BYTE;
	END_VAR

	_BYTE_TO_INT := USINT_TO_INT(BYTE_TO_USINT(IN));
END_FUNCTION

FUNCTION BYTE_OF_DWORD:BYTE
	VAR_INPUT
		IN :	DWORD;
		N :	BYTE;
	END_VAR
	BYTE_OF_DWORD := DWORD_TO_BYTE(SHR(in,_BYTE_TO_INT(SHL(n,3))));
END_FUNCTION

PROGRAM program0
  VAR
    LocalVar0 : DWORD;
	  LocalVar1 : BYTE;
    LocalOUT  : BYTE;
  END_VAR

  LocalOUT := BYTE_OF_DWORD(LocalVar0, LocalVar1);
END_PROGRAM

CONFIGURATION Config0
  RESOURCE Res0 ON PLC
    TASK task0(INTERVAL := T#20ms,PRIORITY := 0);
    PROGRAM instance0 WITH task0 : program0;
  END_RESOURCE
END_CONFIGURATION

(* ---- BYTE_TO_GRAY.ST ---- *)
FUNCTION BYTE_TO_GRAY:BYTE
	VAR_INPUT
		IN :	BYTE;
	END_VAR

	BYTE_TO_GRAY := IN XOR SHR(IN,1);
END_FUNCTION

PROGRAM program0
  VAR
    LocalVar0 : BYTE;
    CEIL5_OUT : BYTE;
  END_VAR

  CEIL5_OUT := BYTE_TO_GRAY(LocalVar0);
END_PROGRAM

CONFIGURATION Config0

  RESOURCE Res0 ON PLC
    TASK task0(INTERVAL := T#20ms,PRIORITY := 0);
    PROGRAM instance0 WITH task0 : program0;
  END_RESOURCE
END_CONFIGURATION

(* ---- BYTE_TO_RANGE.ST ---- *)
FUNCTION _BYTE_TO_REAL:REAL
	VAR_INPUT
		IN :	BYTE;
	END_VAR

	_BYTE_TO_REAL := USINT_TO_REAL(BYTE_TO_USINT(IN));
END_FUNCTION

FUNCTION BYTE_TO_RANGE:REAL
	VAR_INPUT
		X :	BYTE;
		LOW :	REAL;
		HIGH :	REAL;
	END_VAR

	Byte_to_Range := (high - low) * _BYTE_TO_REAL(X) / 255.0 + low;
END_FUNCTION

PROGRAM program0
  VAR
    LocalVar0 : BYTE;
    LocalVar1 : REAL;
	LocalVar2 : REAL;
    CEIL5_OUT : REAL;
  END_VAR

  CEIL5_OUT := BYTE_TO_RANGE(LocalVar0, LocalVar1, LocalVar2);
END_PROGRAM

CONFIGURATION Config0

  RESOURCE Res0 ON PLC
    TASK task0(INTERVAL := T#20ms,PRIORITY := 0);
    PROGRAM instance0 WITH task0 : program0;
  END_RESOURCE
END_CONFIGURATION

(* ---- BYTE_TO_TIME.ST ---- *)
FUNCTION _BYTE_TO_INT:INT
	VAR_INPUT
		IN :	BYTE;
	END_VAR

	_BYTE_TO_INT := USINT_TO_INT(BYTE_TO_USINT(IN));
END_FUNCTION

FUNCTION BYTE_TO_TIME2:TIME
	VAR_INPUT
		IN :	BYTE;
	END_VAR

	BYTE_TO_TIME2 := INT_TO_TIME(_BYTE_TO_INT(IN));
END_FUNCTION

PROGRAM program0
  VAR
    LocalVar0 : BYTE;
    CEIL5_OUT : TIME;
  END_VAR

  CEIL5_OUT := BYTE_TO_TIME2(LocalVar0);
END_PROGRAM

CONFIGURATION Config0

  RESOURCE Res0 ON PLC
    TASK task0(INTERVAL := T#20ms,PRIORITY := 0);
    PROGRAM instance0 WITH task0 : program0;
  END_RESOURCE
END_CONFIGURATION

(* ---- C_TO_F.ST ---- *)
FUNCTION C_TO_F:REAL
	VAR_INPUT
		CELSIUS :	REAL;
	END_VAR

	C_TO_F := celsius * 1.8 + 32.0;
END_FUNCTION

PROGRAM program0
  VAR
    LocalVar0 : REAL;
    CEIL5_OUT : REAL;
  END_VAR

  CEIL5_OUT := C_TO_F(LocalVar0);
END_PROGRAM

CONFIGURATION Config0

  RESOURCE Res0 ON PLC
    TASK task0(INTERVAL := T#20ms,PRIORITY := 0);
    PROGRAM instance0 WITH task0 : program0;
  END_RESOURCE
END_CONFIGURATION

(* ---- C_TO_K.ST ---- *)
FUNCTION C_TO_K:REAL
	VAR_INPUT
		CELSIUS :	REAL;
	END_VAR

	C_to_K := Celsius - 273.15;
END_FUNCTION

PROGRAM program0
  VAR
    LocalVar0 : REAL;
    CEIL5_OUT : REAL;
  END_VAR

  CEIL5_OUT := C_TO_K(LocalVar0);
END_PROGRAM

CONFIGURATION Config0

  RESOURCE Res0 ON PLC
    TASK task0(INTERVAL := T#20ms,PRIORITY := 0);
    PROGRAM instance0 WITH task0 : program0;
  END_RESOURCE
END_CONFIGURATION

(* ---- CAUCHY.ST ---- *)
FUNCTION CAUCHY:REAL
	VAR_INPUT
		X :	REAL;
		T :	REAL;
		U :	REAL;
	END_VAR

	VAR
		tmp :	REAL;
	END_VAR

	tmp := x - t;
	CAUCHY := 0.318309886183791 * U / (U*U + tmp*tmp);
END_FUNCTION

PROGRAM program0
  VAR
    LocalVar0 : REAL;
    LocalVar1 : REAL;
	LocalVar2 : REAL;
    CEIL5_OUT : REAL;
  END_VAR

  CEIL5_OUT := CAUCHY(LocalVar0, LocalVar1, LocalVar2);
END_PROGRAM

CONFIGURATION Config0

  RESOURCE Res0 ON PLC
    TASK task0(INTERVAL := T#20ms,PRIORITY := 0);
    PROGRAM instance0 WITH task0 : program0;
  END_RESOURCE
END_CONFIGURATION

(* ---- CAUCHYCD.ST ---- *)
FUNCTION CAUCHYCD:REAL
	VAR_INPUT
		X :	REAL;
		T :	REAL;
		U :	REAL;
	END_VAR

	CAUCHYCD := 0.5 + 0.318309886183791 * ATAN((X - T) / U);
END_FUNCTION

PROGRAM program0
  VAR
    LocalVar0 : REAL;
	LocalVar1 : REAL;
	LocalVar2 : REAL;
	LocalOUT  : REAL;
  END_VAR
	LocalOUT := CAUCHYCD(LocalVar0, LocalVar1, LocalVar2);
END_PROGRAM

CONFIGURATION Config0
  RESOURCE Res0 ON PLC
    TASK task0(INTERVAL := T#20ms,PRIORITY := 0);
    PROGRAM instance0 WITH task0 : program0;
  END_RESOURCE
END_CONFIGURATION

(* ---- CEIL.ST ---- *)
FUNCTION CEIL:INT

	VAR_INPUT
		X :	REAL;
	END_VAR

	CEIL := REAL_TO_INT(x);
	IF INT_TO_REAL(CEIL) < X THEN
			CEIL := CEIL + 1;
	END_IF;

END_FUNCTION

PROGRAM program0
  VAR
    LocalVar0 : REAL;
    CEIL5_OUT : INT;
  END_VAR

  CEIL5_OUT := CEIL(LocalVar0);
END_PROGRAM

CONFIGURATION Config0

  RESOURCE Res0 ON PLC
    TASK task0(INTERVAL := T#20ms,PRIORITY := 0);
    PROGRAM instance0 WITH task0 : program0;
  END_RESOURCE
END_CONFIGURATION

(* ---- CEIL2.ST ---- *)
FUNCTION _REAL_TO_DINT:DINT
  VAR_INPUT
    X :	REAL;
  END_VAR

  IF REAL_TO_DINT(0.5) = DINT#1 THEN
    _REAL_TO_DINT := REAL_TO_DINT(x);
    RETURN;
  END_IF;

  IF X > 0.0 THEN
    _REAL_TO_DINT := REAL_TO_DINT(x+0.5);
  ELSIF X < 0.0 THEN
    _REAL_TO_DINT := REAL_TO_DINT(x-0.5);
  ELSE
    _REAL_TO_DINT := DINT#0;
  END_IF;
END_FUNCTION

FUNCTION CEIL2:DINT

	VAR_INPUT
		X :	REAL;
	END_VAR

	CEIL2 := _REAL_TO_DINT(x);
	IF DINT_TO_REAL(CEIL2) < X THEN
			CEIL2 := CEIL2 + DINT#1;
	END_IF;

END_FUNCTION

PROGRAM program0
  VAR
    LocalVar0 : REAL;
    CEIL5_OUT : DINT;
  END_VAR

  CEIL5_OUT := CEIL2(LocalVar0);
END_PROGRAM

CONFIGURATION Config0

  RESOURCE Res0 ON PLC
    TASK task0(INTERVAL := T#20ms,PRIORITY := 0);
    PROGRAM instance0 WITH task0 : program0;
  END_RESOURCE
END_CONFIGURATION

(* ---- CHECK_PARITY.ST ---- *)
FUNCTION BIT_OF_DWORD : BOOL
  VAR_INPUT
    IN : DWORD;
    N : INT;
  END_VAR

  BIT_OF_DWORD := (SHR(in,N) AND 16#00000001) > 0;
END_FUNCTION

FUNCTION CHECK_PARITY:BOOL

	VAR_INPUT
		IN :	DWORD;
		P :	BOOL;
	END_VAR

	VAR
		in2 :	DWORD;
	END_VAR

	in2:=in;
	check_parity := NOT p;
	WHILE in2 > DWORD#0 DO
		check_parity := check_parity XOR BIT_OF_DWORD(in2,0) XOR BIT_OF_DWORD(in2,1) XOR BIT_OF_DWORD(in2,2) XOR BIT_OF_DWORD(in2,3);
		in2 := SHR(in2,4);
	END_WHILE;

END_FUNCTION

PROGRAM program0
  VAR
    LocalVar0 : DWORD;
    LocalVar1 : BOOL;
    CEIL5_OUT : BOOL;
  END_VAR

  CEIL5_OUT := CHECK_PARITY(LocalVar0, LocalVar1);
END_PROGRAM

CONFIGURATION Config0

  RESOURCE Res0 ON PLC
    TASK task0(INTERVAL := T#20ms,PRIORITY := 0);
    PROGRAM instance0 WITH task0 : program0;
  END_RESOURCE
END_CONFIGURATION

(* ---- CIRCLE_A.ST ---- *)
FUNCTION CIRCLE_A:REAL
	VAR_INPUT
		RX :	REAL;
		AX :	REAL;
	END_VAR

	circle_A := Rx * RX * 8.726646E-3 * Ax;
END_FUNCTION

PROGRAM program0
  VAR
    LocalVar0 : REAL;
	LocalVar1 : REAL;
	LocalOUT  : REAL;
  END_VAR
  	LocalOUT := CIRCLE_A(LocalVar0, LocalVar1);
END_PROGRAM

CONFIGURATION Config0
  RESOURCE Res0 ON PLC
    TASK task0(INTERVAL := T#20ms,PRIORITY := 0);
    PROGRAM instance0 WITH task0 : program0;
  END_RESOURCE
END_CONFIGURATION

(* ---- CIRCLE_C.ST ---- *)
FUNCTION CIRCLE_C:REAL
	VAR_INPUT
		RX :	REAL;
		AX :	REAL;
	END_VAR

	circle_C := 1.7453293E-2 * Rx * Ax;
END_FUNCTION

PROGRAM program0
  VAR
    LocalVar0 : REAL;
	LocalVar1 : REAL;
	LocalOUT  : REAL;
  END_VAR
  	LocalOUT := CIRCLE_C(LocalVar0, LocalVar1);
END_PROGRAM

CONFIGURATION Config0
  RESOURCE Res0 ON PLC
    TASK task0(INTERVAL := T#20ms,PRIORITY := 0);
    PROGRAM instance0 WITH task0 : program0;
  END_RESOURCE
END_CONFIGURATION

(* ---- CIRCLE_SEG.ST ---- *)
FUNCTION CIRCLE_SEG:REAL
	VAR_INPUT
		RX :	REAL;
		HX :	REAL;
	END_VAR

	IF RX > 0.0 THEN
		CIRCLE_SEG := 2.0 * ACOS(1.0 - LIMIT(0.0, HX / RX, 2.0));
		CIRCLE_SEG := (CIRCLE_SEG - SIN(CIRCLE_SEG)) * RX * RX * 0.5;
	END_IF;
END_FUNCTION

PROGRAM program0
  VAR
    LocalVar0 : REAL;
	LocalVar1 : REAL;
	LocalOUT  : REAL;
  END_VAR
  	LocalOUT := CIRCLE_SEG(LocalVar0, LocalVar1);
END_PROGRAM

CONFIGURATION Config0
  RESOURCE Res0 ON PLC
    TASK task0(INTERVAL := T#20ms,PRIORITY := 0);
    PROGRAM instance0 WITH task0 : program0;
  END_RESOURCE
END_CONFIGURATION

(* ---- CMP.ST ---- *)
FUNCTION EXP10 : REAL
  VAR_INPUT
    x : REAL;
  END_VAR

  exp10 := EXP(X * 2.30258509299405);
  (* from OSCAT library; www.oscat.de  *)
END_FUNCTION

FUNCTION FLOOR : INT
  VAR_INPUT
    x : REAL;
  END_VAR

  FLOOR := REAL_TO_INT(X);
  IF INT_TO_REAL(FLOOR) > X THEN
  	floor := floor - 1;
  END_IF;
  (* from OSCAT library; www.oscat.de  *)
END_FUNCTION

FUNCTION CMP:BOOL
	VAR_INPUT
		X :	REAL;
		Y :	REAL;
		N :	INT;
	END_VAR

	VAR
		tmp :	REAL;
	END_VAR

	tmp := ABS(x);
	IF tmp > 0.0 THEN
		tmp := EXP10(INT_TO_REAL(FLOOR(LOG(tmp))-N+1));
	ELSE
		tmp := EXP10(tmp);
	END_IF;
	CMP := ABS(X - Y) < tmp;

END_FUNCTION

PROGRAM program0
  VAR
    LocalVar0 : REAL;
    LocalVar1 : REAL;
	LocalVar2 : INT;
    CEIL5_OUT : BOOL;
  END_VAR

  CEIL5_OUT := CMP(LocalVar0, LocalVar1, LocalVar2);
END_PROGRAM

CONFIGURATION Config0

  RESOURCE Res0 ON PLC
    TASK task0(INTERVAL := T#20ms,PRIORITY := 0);
    PROGRAM instance0 WITH task0 : program0;
  END_RESOURCE
END_CONFIGURATION

(* ---- CONE_V.ST ---- *)
FUNCTION CONE_V:REAL
	VAR_INPUT
		RX :	REAL;
		HX :	REAL;
	END_VAR

	cone_V := 1.047197551 * RX * RX * hx;
END_FUNCTION

PROGRAM program0
  VAR
    LocalVar0 : REAL;
	LocalVar1 : REAL;
	LocalOUT  : REAL;
  END_VAR
  	LocalOUT := CONE_V(LocalVar0, LocalVar1);
END_PROGRAM

CONFIGURATION Config0
  RESOURCE Res0 ON PLC
    TASK task0(INTERVAL := T#20ms,PRIORITY := 0);
    PROGRAM instance0 WITH task0 : program0;
  END_RESOURCE
END_CONFIGURATION

(* ---- COSH.ST ---- *)
FUNCTION COSH:REAL
	VAR_INPUT
		X :	REAL;
	END_VAR

	VAR
		t :	REAL;
	END_VAR

	T := EXP(X);
	COSH := (1.0 / T + T) * 0.5;
END_FUNCTION

PROGRAM program0
  VAR
    LocalVar0 : REAL;
    CEIL5_OUT : REAL;
  END_VAR

  CEIL5_OUT := COSH(LocalVar0);
END_PROGRAM

CONFIGURATION Config0

  RESOURCE Res0 ON PLC
    TASK task0(INTERVAL := T#20ms,PRIORITY := 0);
    PROGRAM instance0 WITH task0 : program0;
  END_RESOURCE
END_CONFIGURATION

(* ---- COTH.ST ---- *)
FUNCTION COTH:REAL

	VAR_INPUT
		X :	REAL;
	END_VAR

	IF X > 20.0 THEN
		COTH :=1.0;
	ELSIF X < -20.0 THEN
		COTH := -1.0;
	ELSE
		COTH := 1.0 + 2.0 / (EXP(X * 2.0) - 1.0);
	END_IF;

END_FUNCTION

PROGRAM program0
	VAR
		X :	REAL;
		OUT : REAL;
	END_VAR

	OUT := COTH(X);

END_PROGRAM

CONFIGURATION Config0

	RESOURCE Res0 ON PLC
		TASK task0(INTERVAL := T#20ms,PRIORITY := 0);
		PROGRAM instance0 WITH task0 : program0;
	END_RESOURCE

END_CONFIGURATION

(* ---- CTRL_IN.ST ---- *)
FUNCTION DEAD_ZONE:REAL

	VAR_INPUT
		X :	REAL;
		L :	REAL;
	END_VAR

	IF ABS(x) > L THEN
		dead_zone := X;
	ELSE
		DEAD_ZONE := 0.0;
	END_IF;

END_FUNCTION

FUNCTION CTRL_IN:REAL
	VAR_INPUT
		SET_POINT :	REAL;
		ACTUAL :	REAL;
		NOISE :	REAL;
	END_VAR
	CTRL_IN := DEAD_ZONE(SET_POINT - ACTUAL, NOISE);
END_FUNCTION

PROGRAM program0
  VAR
    LocalVar0 : REAL;
	LocalVar1 : REAL;
	LocalVar2 : REAL;
	LocalOUT  : REAL;
  END_VAR
  	LocalOUT := CTRL_IN(LocalVar0, LocalVar1, LocalVar2);
END_PROGRAM

CONFIGURATION Config0
  RESOURCE Res0 ON PLC
    TASK task0(INTERVAL := T#20ms,PRIORITY := 0);
    PROGRAM instance0 WITH task0 : program0;
  END_RESOURCE
END_CONFIGURATION

(* ---- D_TRUNC.ST ---- *)
FUNCTION D_TRUNC : DINT
  VAR_INPUT
    x : REAL;
  END_VAR

  D_TRUNC := REAL_TO_DINT(X);
  IF X > 0.0 THEN
  	IF DINT_TO_REAL(D_TRUNC) > X THEN D_TRUNC := D_TRUNC - DINT#1; END_IF;
  ELSE
  	IF DINT_TO_REAL(D_TRUNC) < X THEN D_TRUNC := D_TRUNC + DINT#1; END_IF;
  END_IF;
END_FUNCTION

PROGRAM program0
  VAR
    LocalVar0 : REAL;
    LocalVar1 : DINT;
    CEIL5_OUT : DINT;
  END_VAR

  CEIL5_OUT := D_TRUNC(LocalVar0);
  LocalVar1 := CEIL5_OUT;
END_PROGRAM

CONFIGURATION Config0

  RESOURCE Res0 ON PLC
    TASK task0(INTERVAL := T#20ms,PRIORITY := 0);
    PROGRAM instance0 WITH task0 : program0;
  END_RESOURCE
END_CONFIGURATION

(* ---- DATE_ADD.ST ---- *)
FUNCTION YEAR_OF_DATE:INT
	VAR_INPUT
		IDATE :	UDINT;
	END_VAR

	YEAR_OF_DATE := UDINT_TO_INT((idate+UDINT#43200) / UDINT#31557600 + UDINT#1970);
END_FUNCTION

FUNCTION DAY_OF_WEEK:INT

	VAR_INPUT
		IDATE :	UDINT;
	END_VAR

	DAY_OF_WEEK := UDINT_TO_INT((idate / UDINT#86400 + UDINT#3) MOD UDINT#7) + INT#01;
END_FUNCTION

FUNCTION LEAP_OF_DATE:BOOL

	VAR_INPUT
		IDATE :	UDINT;
	END_VAR

	LEAP_OF_DATE := SHL(UDINT_TO_DWORD((idate + UDINT#43200) / UDINT#31557600), 30) = DWORD#16#80000000;
END_FUNCTION

FUNCTION DAY_OF_YEAR:INT
	VAR_INPUT
		IDATE :	UDINT;
	END_VAR

	DAY_OF_YEAR := UDINT_TO_INT(((idate) / UDINT#86400) MOD UDINT#1461);
	IF DAY_OF_YEAR > 729 THEN
		IF DAY_OF_YEAR > 1095 THEN DAY_OF_YEAR := DAY_OF_YEAR - 1095; ELSE DAY_OF_YEAR := DAY_OF_YEAR - 729; END_IF;
	ELSIF DAY_OF_YEAR > 364 THEN
		DAY_OF_YEAR := DAY_OF_YEAR - 364;
	ELSE
		DAY_OF_YEAR := DAY_OF_YEAR + 1;
	END_IF;
END_FUNCTION

FUNCTION MONTH_OF_DATE:INT

	VAR_INPUT
		IDATE :	UDINT;
	END_VAR

	MONTH_OF_DATE := DAY_OF_YEAR(idate);
	IF MONTH_OF_DATE < 32 THEN
		MONTH_OF_DATE := 1;
	ELSIF LEAP_OF_DATE((IDATE)) THEN
		MONTH_OF_DATE := (MONTH_OF_DATE * 53 + 1668) / 1623;
	ELSE
		MONTH_OF_DATE := (MONTH_OF_DATE * 53 + 1700) / 1620;
	END_IF;
END_FUNCTION

FUNCTION DAY_OF_MONTH:INT
	VAR_INPUT
		IDATE :	UDINT;
	END_VAR

	day_of_month := day_of_year(idate);

	IF leap_of_Date((idate)) THEN
		CASE day_of_month OF
			32..60	:	day_of_month := day_of_month - 31;
			61..91	:	day_of_month := day_of_month - 60;
			92..121 :	day_of_month := day_of_month - 91;
			122..152:	day_of_month := day_of_month - 121;
			153..182:	day_of_month := day_of_month - 152;
			183..213:	day_of_month := day_of_month - 182;
			214..244:	day_of_month := day_of_month - 213;
			245..274:	day_of_month := day_of_month - 244;
			275..305:	day_of_month := day_of_month - 274;
			306..335:	day_of_month := day_of_month - 305;
			336..366:	day_of_month := day_of_month - 335;
		END_CASE;
	ELSE
		CASE day_of_month OF
			32..59	:	day_of_month := day_of_month - 31;
			60..90	:	day_of_month := day_of_month - 59;
			91..120 :	day_of_month := day_of_month - 90;
			121..151:	day_of_month := day_of_month - 120;
			152..181:	day_of_month := day_of_month - 151;
			182..212:	day_of_month := day_of_month - 181;
			213..243:	day_of_month := day_of_month - 212;
			244..273:	day_of_month := day_of_month - 243;
			274..304:	day_of_month := day_of_month - 273;
			305..334:	day_of_month := day_of_month - 304;
			335..365:	day_of_month := day_of_month - 334;
		END_CASE;
	END_IF;
END_FUNCTION

FUNCTION _INT_TO_UDINT:UDINT
	VAR_INPUT
		IN :	INT;
	END_VAR

	_INT_TO_UDINT := DINT_TO_UDINT(INT_TO_DINT(IN));
END_FUNCTION

FUNCTION SET_DATE:UDINT

	VAR_INPUT
		YEAR :	INT;
		MONTH :	INT;
		DAY :	INT;
	END_VAR

	VAR
		count :	INT;
	END_VAR

	IF month > 2 THEN
		count := (month - 1) * 30;
		IF month > 7 THEN
			count := count + DWORD_TO_INT(SHR(DINT_TO_DWORD(INT_TO_DINT(month) - INT_TO_DINT(3)),1));
		ELSE
			count := count + DWORD_TO_INT(SHR(DINT_TO_DWORD(INT_TO_DINT(month) - INT_TO_DINT(4)),1));
		END_IF;
		IF SHL(INT_TO_WORD(year),14) = WORD#0 THEN
			count := count + 1;
		END_IF;
	ELSE
		count := (month - 1) * 31;
	END_IF;
	SET_DATE := (_INT_TO_UDINT(count + day - 1) + DWORD_TO_UDINT(SHR(UDINT_TO_DWORD(_INT_TO_UDINT(year) * UDINT#1461 - UDINT#2878169), 2))) * UDINT#86400;

END_FUNCTION

FUNCTION DATE_ADD:UDINT
	VAR_INPUT
		IDATE :	UDINT;
		D :	INT;
		W :	INT;
		M :	INT;
		Y :	INT;
	END_VAR

	VAR
		mo :	INT;
		yr :	INT;
		dm :	INT;
	END_VAR

	DATE_ADD := IDATE + INT_TO_UDINT(D + W * 7) * UDINT#86400;
	yr := Y + YEAR_OF_DATE(DATE_ADD);
	mo := M + MONTH_OF_DATE(DATE_ADD);
	dm := DAY_OF_MONTH(DATE_ADD);
	WHILE mo > 12 DO
		mo := mo - 12;
		yr := yr + 1;
	END_WHILE;
	WHILE mo < 1 DO
		mo := mo + 12;
		yr := yr - 1;
	END_WHILE;
	DATE_ADD := SET_DATE(yr, mo, dm);
END_FUNCTION

PROGRAM program0
  VAR
    LocalVar0 : UDINT;
	LocalVar1 : INT;
	LocalVar2 : INT;
	LocalVar3 : INT;
	LocalVar4 : INT;
	LocalOUT  : UDINT;
  END_VAR
  	LocalOUT := DATE_ADD(LocalVar0, LocalVar1, LocalVar2, LocalVar3, LocalVar4);
END_PROGRAM

CONFIGURATION Config0
  RESOURCE Res0 ON PLC
    TASK task0(INTERVAL := T#20ms,PRIORITY := 0);
    PROGRAM instance0 WITH task0 : program0;
  END_RESOURCE
END_CONFIGURATION

(* ---- DATE_TO_DT.ST ---- *)
FUNCTION DATE_TO_DT:UDINT
	VAR_INPUT
		IN :	UDINT;
	END_VAR
	DATE_TO_DT := IN;
END_FUNCTION

PROGRAM program0
  VAR
    LocalVar0 : UDINT;
	LocalOUT  : UDINT;
  END_VAR
  	LocalOUT := DATE_TO_DT(LocalVar0);
END_PROGRAM

CONFIGURATION Config0
  RESOURCE Res0 ON PLC
    TASK task0(INTERVAL := T#20ms,PRIORITY := 0);
    PROGRAM instance0 WITH task0 : program0;
  END_RESOURCE
END_CONFIGURATION

(* ---- DATE_TO_DWORD.ST ---- *)
FUNCTION DATE_TO_DWORD2:DWORD
	VAR_INPUT
		IN :	UDINT;
	END_VAR

	DATE_TO_DWORD2 := UDINT_TO_DWORD(IN);
END_FUNCTION

PROGRAM program0
  VAR
    LocalVar0 : UDINT;
	LocalOUT  : DWORD;
  END_VAR
  	LocalOUT := DATE_TO_DWORD2(LocalVar0);
END_PROGRAM

CONFIGURATION Config0
  RESOURCE Res0 ON PLC
    TASK task0(INTERVAL := T#20ms,PRIORITY := 0);
    PROGRAM instance0 WITH task0 : program0;
  END_RESOURCE
END_CONFIGURATION

(* ---- DATE_TO_REAL.ST ---- *)
FUNCTION DATE_TO_REAL2:REAL
	VAR_INPUT
		IN :	UDINT;
	END_VAR

	DATE_TO_REAL2 := UDINT_TO_REAL(IN);
END_FUNCTION

PROGRAM program0
  VAR
    LocalVar0 : UDINT;
	LocalOUT  : REAL;
  END_VAR
  	LocalOUT := DATE_TO_REAL2(LocalVar0);
END_PROGRAM

CONFIGURATION Config0
  RESOURCE Res0 ON PLC
    TASK task0(INTERVAL := T#20ms,PRIORITY := 0);
    PROGRAM instance0 WITH task0 : program0;
  END_RESOURCE
END_CONFIGURATION

(* ---- DATE_TO_UDINT.ST ---- *)
FUNCTION DATE_TO_UDINT2:UDINT
	VAR_INPUT
		IN :	UDINT;
	END_VAR

	DATE_TO_UDINT2 := IN;
END_FUNCTION

PROGRAM program0
  VAR
    LocalVar0 : UDINT;
	LocalOUT  : UDINT;
  END_VAR
  	LocalOUT := DATE_TO_UDINT2(LocalVar0);
END_PROGRAM

CONFIGURATION Config0
  RESOURCE Res0 ON PLC
    TASK task0(INTERVAL := T#20ms,PRIORITY := 0);
    PROGRAM instance0 WITH task0 : program0;
  END_RESOURCE
END_CONFIGURATION

(* ---- DAY_OF_DATE.ST ---- *)
FUNCTION DAY_OF_DATE:DINT
	VAR_INPUT
		IDATE :	UDINT;
	END_VAR

	day_of_date := UDINT_TO_DINT(idate / UDINT#86400);
END_FUNCTION

PROGRAM program0
  VAR
    LocalVar0 : UDINT;
	LocalOUT  : DINT;
  END_VAR
  	LocalOUT := DAY_OF_DATE(LocalVar0);
END_PROGRAM

CONFIGURATION Config0
  RESOURCE Res0 ON PLC
    TASK task0(INTERVAL := T#20ms,PRIORITY := 0);
    PROGRAM instance0 WITH task0 : program0;
  END_RESOURCE
END_CONFIGURATION

(* ---- DAY_OF_MONTH.ST ---- *)
FUNCTION LEAP_OF_DATE:BOOL

	VAR_INPUT
		IDATE :	UDINT;
	END_VAR

	LEAP_OF_DATE := SHL(UDINT_TO_DWORD((idate + UDINT#43200) / UDINT#31557600), 30) = DWORD#16#80000000;

END_FUNCTION

FUNCTION DAY_OF_YEAR:INT
	VAR_INPUT
		IDATE :	DATE;
	END_VAR

	DAY_OF_YEAR := UDINT_TO_INT((DATE_TO_UDINT(idate) / UDINT#86400) MOD UDINT#1461);
	IF DAY_OF_YEAR > 729 THEN
		IF DAY_OF_YEAR > 1095 THEN DAY_OF_YEAR := DAY_OF_YEAR - 1095; ELSE DAY_OF_YEAR := DAY_OF_YEAR - 729; END_IF;
	ELSIF DAY_OF_YEAR > 364 THEN
		DAY_OF_YEAR := DAY_OF_YEAR - 364;
	ELSE
		DAY_OF_YEAR := DAY_OF_YEAR + 1;
	END_IF;
END_FUNCTION

FUNCTION DAY_OF_MONTH:INT
	VAR_INPUT
		IDATE :	DATE;
	END_VAR

	day_of_month := day_of_year(idate);

	IF leap_of_Date(DATE_TO_UDINT(idate)) THEN
		CASE day_of_month OF
			32..60	:	day_of_month := day_of_month - 31;
			61..91	:	day_of_month := day_of_month - 60;
			92..121 :	day_of_month := day_of_month - 91;
			122..152:	day_of_month := day_of_month - 121;
			153..182:	day_of_month := day_of_month - 152;
			183..213:	day_of_month := day_of_month - 182;
			214..244:	day_of_month := day_of_month - 213;
			245..274:	day_of_month := day_of_month - 244;
			275..305:	day_of_month := day_of_month - 274;
			306..335:	day_of_month := day_of_month - 305;
			336..366:	day_of_month := day_of_month - 335;
		END_CASE;
	ELSE
		CASE day_of_month OF
			32..59	:	day_of_month := day_of_month - 31;
			60..90	:	day_of_month := day_of_month - 59;
			91..120 :	day_of_month := day_of_month - 90;
			121..151:	day_of_month := day_of_month - 120;
			152..181:	day_of_month := day_of_month - 151;
			182..212:	day_of_month := day_of_month - 181;
			213..243:	day_of_month := day_of_month - 212;
			244..273:	day_of_month := day_of_month - 243;
			274..304:	day_of_month := day_of_month - 273;
			305..334:	day_of_month := day_of_month - 304;
			335..365:	day_of_month := day_of_month - 334;
		END_CASE;
	END_IF;

END_FUNCTION

PROGRAM program0
  VAR
    LocalVar0 : DATE;
	LocalOUT  : INT;
  END_VAR
  	LocalOUT := DAY_OF_MONTH(LocalVar0);
END_PROGRAM

CONFIGURATION Config0
  RESOURCE Res0 ON PLC
    TASK task0(INTERVAL := T#20ms,PRIORITY := 0);
    PROGRAM instance0 WITH task0 : program0;
  END_RESOURCE
END_CONFIGURATION

(* ---- DAY_OF_WEEK.ST ---- *)
FUNCTION DAY_OF_WEEK:INT
  VAR_INPUT
    IDATE :	UDINT;
  END_VAR

  DAY_OF_WEEK := UDINT_TO_INT((idate / UDINT#86400 + UDINT#3) MOD UDINT#7) + INT#01;
END_FUNCTION

PROGRAM program0
  VAR
    LocalVar0 : UDINT;
	LocalOUT  : INT;
  END_VAR
  	LocalOUT := DAY_OF_WEEK(LocalVar0);
END_PROGRAM

CONFIGURATION Config0
  RESOURCE Res0 ON PLC
    TASK task0(INTERVAL := T#20ms,PRIORITY := 0);
    PROGRAM instance0 WITH task0 : program0;
  END_RESOURCE
END_CONFIGURATION

(* ---- DAY_OF_YEAR.ST ---- *)
FUNCTION DAY_OF_YEAR:INT
	VAR_INPUT
		IDATE :	DATE;
	END_VAR

	DAY_OF_YEAR := UDINT_TO_INT((DATE_TO_UDINT(idate) / UDINT#86400) MOD UDINT#1461);
	IF DAY_OF_YEAR > 729 THEN
		IF DAY_OF_YEAR > 1095 THEN DAY_OF_YEAR := DAY_OF_YEAR - 1095; ELSE DAY_OF_YEAR := DAY_OF_YEAR - 729; END_IF;
	ELSIF DAY_OF_YEAR > 364 THEN
		DAY_OF_YEAR := DAY_OF_YEAR - 364;
	ELSE
		DAY_OF_YEAR := DAY_OF_YEAR + 1;
	END_IF;
END_FUNCTION

PROGRAM program0
  VAR
    LocalVar0 : DATE;
	LocalOUT  : INT;
  END_VAR
  	LocalOUT := DAY_OF_YEAR(LocalVar0);
END_PROGRAM

CONFIGURATION Config0
  RESOURCE Res0 ON PLC
    TASK task0(INTERVAL := T#20ms,PRIORITY := 0);
    PROGRAM instance0 WITH task0 : program0;
  END_RESOURCE
END_CONFIGURATION

(* ---- DAY_TO_TIME.ST ---- *)
FUNCTION DAY_TO_TIME:TIME
	VAR_INPUT
		IN :	REAL;
	END_VAR

	day_to_time := DINT_TO_TIME(UDINT_TO_DINT(_REAL_TO_UDINT(IN * REAL#86400000.00)));
END_FUNCTION

FUNCTION _REAL_TO_UDINT:UDINT
  VAR_INPUT
    X :	REAL;
  END_VAR

  IF REAL_TO_UDINT(0.5) = UDINT#1 THEN
    _REAL_TO_UDINT := REAL_TO_UDINT(x);
  ELSIF X > 0.0 THEN
    _REAL_TO_UDINT := REAL_TO_UDINT(x+0.5);
  ELSIF X < 0.0 THEN
    _REAL_TO_UDINT := REAL_TO_UDINT(x-0.5);
  ELSE
    _REAL_TO_UDINT := UDINT#0;
  END_IF;
END_FUNCTION

PROGRAM program0
  VAR
    LocalVar0 : REAL;
	LocalOUT  : TIME;
  END_VAR
  	LocalOUT := DAY_TO_TIME(LocalVar0);
END_PROGRAM

CONFIGURATION Config0
  RESOURCE Res0 ON PLC
    TASK task0(INTERVAL := T#20ms,PRIORITY := 0);
    PROGRAM instance0 WITH task0 : program0;
  END_RESOURCE
END_CONFIGURATION

(* ---- DAYS_DELTA.ST ---- *)
FUNCTION DAYS_DELTA:DINT
	VAR_INPUT
		DATE_1 :	UDINT;
		DATE_2 :	UDINT;
	END_VAR
	IF DATE_1 > DATE_2 THEN
		DAYS_DELTA := - UDINT_TO_DINT((date_1 - date_2) / UDINT#86400);
	ELSE
		DAYS_DELTA :=   UDINT_TO_DINT((date_2 - date_1) / UDINT#86400);
	END_IF;
END_FUNCTION

PROGRAM program0
  VAR
    LocalVar0 : UDINT;
	LocalVar1 : UDINT;
	LocalOUT  : DINT;
  END_VAR
  	LocalOUT := DAYS_DELTA(LocalVar0, LocalVar1);
END_PROGRAM

CONFIGURATION Config0
  RESOURCE Res0 ON PLC
    TASK task0(INTERVAL := T#20ms,PRIORITY := 0);
    PROGRAM instance0 WITH task0 : program0;
  END_RESOURCE
END_CONFIGURATION

(* ---- DAYS_IN_MONTH.ST ---- *)
FUNCTION DAY_OF_YEAR:INT
	VAR_INPUT
		IDATE :	UDINT;
	END_VAR

	DAY_OF_YEAR := UDINT_TO_INT(((idate) / UDINT#86400) MOD UDINT#1461);
	IF DAY_OF_YEAR > 729 THEN
		IF DAY_OF_YEAR > 1095 THEN DAY_OF_YEAR := DAY_OF_YEAR - 1095; ELSE DAY_OF_YEAR := DAY_OF_YEAR - 729; END_IF;
	ELSIF DAY_OF_YEAR > 364 THEN
		DAY_OF_YEAR := DAY_OF_YEAR - 364;
	ELSE
		DAY_OF_YEAR := DAY_OF_YEAR + 1;
	END_IF;
END_FUNCTION

FUNCTION LEAP_OF_DATE:BOOL

	VAR_INPUT
		IDATE :	UDINT;
	END_VAR

	LEAP_OF_DATE := SHL(UDINT_TO_DWORD((idate + UDINT#43200) / UDINT#31557600), 30) = DWORD#16#80000000;
END_FUNCTION

FUNCTION DAYS_IN_MONTH:INT

	VAR_INPUT
		IDATE :	UDINT;
	END_VAR

	DAYS_IN_MONTH := DAY_OF_YEAR(IDATE);
	IF LEAP_OF_DATE(IDATE) THEN
		CASE DAYS_IN_MONTH OF
			32..60	:	DAYS_IN_MONTH := 29;
			92..121 :	DAYS_IN_MONTH := 30;
			153..182:	DAYS_IN_MONTH := 30;
			245..274:	DAYS_IN_MONTH := 30;
			306..335:	DAYS_IN_MONTH := 30;
		ELSE
			DAYS_IN_MONTH := 31;
		END_CASE;
	ELSE
		CASE DAYS_IN_MONTH OF
			32..59	:	DAYS_IN_MONTH := 28;
			91..120 :	DAYS_IN_MONTH := 30;
			152..181:	DAYS_IN_MONTH := 30;
			244..273:	DAYS_IN_MONTH := 30;
			305..334:	DAYS_IN_MONTH := 30;
		ELSE
			DAYS_IN_MONTH := 31;
		END_CASE;
	END_IF;

END_FUNCTION

PROGRAM program0
  VAR
    LocalVar0 : UDINT;
	LocalOUT  : INT;
  END_VAR
  	LocalOUT := DAYS_IN_MONTH(LocalVar0);
END_PROGRAM

CONFIGURATION Config0
  RESOURCE Res0 ON PLC
    TASK task0(INTERVAL := T#20ms,PRIORITY := 0);
    PROGRAM instance0 WITH task0 : program0;
  END_RESOURCE
END_CONFIGURATION

(* ---- DAYS_IN_YEAR.ST ---- *)
FUNCTION LEAP_OF_DATE:BOOL

	VAR_INPUT
		IDATE :	UDINT;
	END_VAR

	LEAP_OF_DATE := SHL(UDINT_TO_DWORD((idate + UDINT#43200) / UDINT#31557600), 30) = DWORD#16#80000000;
END_FUNCTION

FUNCTION DAYS_IN_YEAR:INT
	VAR_INPUT
		IDATE :	UDINT;
	END_VAR

	IF LEAP_OF_DATE(IDATE) THEN
		DAYS_IN_YEAR := 366;
	ELSE
		DAYS_IN_YEAR := 365;
	END_IF;
END_FUNCTION

PROGRAM program0
  VAR
    LocalVar0 : UDINT;
	LocalOUT  : INT;
  END_VAR
  	LocalOUT := DAYS_IN_YEAR(LocalVar0);
END_PROGRAM

CONFIGURATION Config0
  RESOURCE Res0 ON PLC
    TASK task0(INTERVAL := T#20ms,PRIORITY := 0);
    PROGRAM instance0 WITH task0 : program0;
  END_RESOURCE
END_CONFIGURATION

(* ---- DEAD_BAND.ST ---- *)
FUNCTION DEAD_BAND:REAL

	VAR_INPUT
		X :	REAL;
		L :	REAL;
	END_VAR

	IF X > L THEN
		DEAD_BAND := X - L;
	ELSIF X < -L THEN
		DEAD_BAND := X + L;
	ELSE
		DEAD_BAND := 0.0;
	END_IF;

END_FUNCTION

PROGRAM program0
  VAR
    LocalVar0 : REAL;
	LocalVar1 : REAL;
	LocalOUT  : REAL;
  END_VAR
  	LocalOUT := DEAD_BAND(LocalVar0, LocalVar1);
END_PROGRAM

CONFIGURATION Config0
  RESOURCE Res0 ON PLC
    TASK task0(INTERVAL := T#20ms,PRIORITY := 0);
    PROGRAM instance0 WITH task0 : program0;
  END_RESOURCE
END_CONFIGURATION

(* ---- DEAD_ZONE.ST ---- *)
FUNCTION DEAD_ZONE:REAL

	VAR_INPUT
		X :	REAL;
		L :	REAL;
	END_VAR

	IF ABS(x) > L THEN
		dead_zone := X;
	ELSE
		DEAD_ZONE := 0.0;
	END_IF;

END_FUNCTION

PROGRAM program0
  VAR
    LocalVar0 : REAL;
	LocalVar1 : REAL;
	LocalOUT  : REAL;
  END_VAR
  	LocalOUT := DEAD_ZONE(LocalVar0, LocalVar1);
END_PROGRAM

CONFIGURATION Config0
  RESOURCE Res0 ON PLC
    TASK task0(INTERVAL := T#20ms,PRIORITY := 0);
    PROGRAM instance0 WITH task0 : program0;
  END_RESOURCE
END_CONFIGURATION

(* ---- DEC1.ST ---- *)
FUNCTION DEC1:INT

	VAR_INPUT
		X :	INT;
		N :	INT;
	END_VAR

	IF X = 0 THEN
		DEC1 := N - 1;
	ELSE
		DEC1 := X - 1;
	END_IF;

END_FUNCTION

PROGRAM program0
  VAR
    LocalVar0 : INT;
	LocalVar1 : INT;
	LocalOUT  : INT;
  END_VAR
  	LocalOUT := DEC1(LocalVar0, LocalVar1);
END_PROGRAM

CONFIGURATION Config0
  RESOURCE Res0 ON PLC
    TASK task0(INTERVAL := T#20ms,PRIORITY := 0);
    PROGRAM instance0 WITH task0 : program0;
  END_RESOURCE
END_CONFIGURATION

(* ---- DEG.ST ---- *)
FUNCTION FLOOR2 : DINT
	VAR_INPUT
		x : REAL;
	END_VAR

	FLOOR2 := REAL_TO_DINT(X);
	IF DINT_TO_REAL(FLOOR2) > X THEN
		FLOOR2 := FLOOR2 - DINT#1;
	END_IF;

END_FUNCTION

FUNCTION MODR:REAL

	VAR_INPUT
		IN :	REAL;
		DIVI :	REAL;
	END_VAR

	IF divi = 0.0 THEN
		MODR := 0.0;
	ELSE
		MODR := in - DINT_TO_REAL(FLOOR2(in / divi)) * divi;
	END_IF;

END_FUNCTION

FUNCTION DEG:REAL

	VAR_INPUT
		RAD :	REAL;
	END_VAR

	DEG := MODR(57.29577951308232 * RAD, 360.0);

END_FUNCTION

PROGRAM program0

	VAR
		RAD :	REAL;
		CEIL5_OUT : REAL;
	END_VAR

	CEIL5_OUT := DEG(RAD);

END_PROGRAM

CONFIGURATION Config0

	RESOURCE Res0 ON PLC
		TASK task0(INTERVAL := T#20ms,PRIORITY := 0);
		PROGRAM instance0 WITH task0 : program0;
	END_RESOURCE

END_CONFIGURATION

(* ---- DEW_CON.ST ---- *)
FUNCTION SDD:REAL

	VAR_INPUT
		T :	REAL;
		ICE :	BOOL;
	END_VAR

	IF ice THEN
		SDD := 611.153 * EXP(22.4433 * T / (272.186 + T));
	ELSE
		SDD := 611.213 * EXP(17.5043 * T / (241.2 + T));
	END_IF;

END_FUNCTION

FUNCTION DEW_CON:REAL

	VAR_INPUT
		RH :	REAL;
		T :	REAL;
	END_VAR

	IF RH > 0.0 AND T > -50.0 THEN
		DEW_CON := 2.166824303E-2 * RH * SDD(T,FALSE)  / (T - -273.15);
	ELSE
		DEW_CON := 0.0;
	END_IF;

END_FUNCTION

PROGRAM program0
  VAR
    RH :	REAL;
	T :	REAL;
    CEIL5_OUT : REAL;
  END_VAR

  CEIL5_OUT := DEW_CON(RH, T);
END_PROGRAM

CONFIGURATION Config0

  RESOURCE Res0 ON PLC
    TASK task0(INTERVAL := T#20ms,PRIORITY := 0);
    PROGRAM instance0 WITH task0 : program0;
  END_RESOURCE
END_CONFIGURATION

(* ---- DEW_RH.ST ---- *)
FUNCTION SDD:REAL

	VAR_INPUT
		T :	REAL;
		ICE :	BOOL;
	END_VAR

	IF ice THEN
		SDD := 611.153 * EXP(22.4433 * T / (272.186 + T));
	ELSE
		SDD := 611.213 * EXP(17.5043 * T / (241.2 + T));
	END_IF;

END_FUNCTION

FUNCTION DEW_CON:REAL

	VAR_INPUT
		RH :	REAL;
		T :	REAL;
	END_VAR

	IF RH > 0.0 AND T > -50.0 THEN
		DEW_CON := 2.166824303E-2 * RH * SDD(T,FALSE)  / (T - -273.15);
	ELSE
		DEW_CON := 0.0;
	END_IF;

END_FUNCTION

FUNCTION DEW_RH:REAL

	VAR_INPUT
		VC :	REAL;
		T :	REAL;
	END_VAR

	DEW_RH := LIMIT(0.0, VC / DEW_CON(1.0, T), 100.0);

END_FUNCTION

PROGRAM program0
	VAR
		VC :	REAL;
		T :	REAL;
		CEIL5_OUT : REAL;
	END_VAR

  	CEIL5_OUT := DEW_RH(VC, T);
END_PROGRAM

CONFIGURATION Config0

  RESOURCE Res0 ON PLC
    TASK task0(INTERVAL := T#20ms,PRIORITY := 0);
    PROGRAM instance0 WITH task0 : program0;
  END_RESOURCE
END_CONFIGURATION

(* ---- DEW_TEMP.ST ---- *)
FUNCTION EXP10 : REAL
  VAR_INPUT
    x : REAL;
  END_VAR

  exp10 := EXP(X * 2.30258509299405);
  (* from OSCAT library; www.oscat.de  *)
END_FUNCTION

FUNCTION DEW_TEMP:REAL

VAR_INPUT
	RH :	REAL;
	T :	REAL;
END_VAR

	VAR
		V :	REAL;
	END_VAR

	IF rh > 0.0 THEN

		V := LOG(RH * 0.01 * EXP10((7.5*T) / (237.3+T)));
		DEW_TEMP := 237.3*V / (7.5-V);
	ELSE
		DEW_TEMP:= -273.15;
	END_IF;

END_FUNCTION

PROGRAM program0
	VAR
		RH :	REAL;
		T :	REAL;
		CEIL5_OUT : REAL;
	END_VAR

  	CEIL5_OUT := DEW_TEMP(RH, T);
END_PROGRAM

CONFIGURATION Config0

  RESOURCE Res0 ON PLC
    TASK task0(INTERVAL := T#20ms,PRIORITY := 0);
    PROGRAM instance0 WITH task0 : program0;
  END_RESOURCE
END_CONFIGURATION

(* ---- DIFFER.ST ---- *)
FUNCTION DIFFER:BOOL
	VAR_INPUT
		IN1 :	REAL;
		IN2 :	REAL;
		X :	REAL;
	END_VAR

	DIFFER := ABS(in1 - in2) > X;
END_FUNCTION

PROGRAM program0
  VAR
    LocalVar0 : REAL;
	LocalVar1 : REAL;
	LocalVar2 : REAL;
	LocalOUT  : BOOL;
  END_VAR
  	LocalOUT := DIFFER(LocalVar0, LocalVar1, LocalVar2);
END_PROGRAM

CONFIGURATION Config0
  RESOURCE Res0 ON PLC
    TASK task0(INTERVAL := T#20ms,PRIORITY := 0);
    PROGRAM instance0 WITH task0 : program0;
  END_RESOURCE
END_CONFIGURATION

(* ---- DST.ST ---- *)
FUNCTION _INT_TO_UDINT:UDINT
	VAR_INPUT
		IN :	INT;
	END_VAR

	_INT_TO_UDINT := DINT_TO_UDINT(INT_TO_DINT(IN));
END_FUNCTION

FUNCTION YEAR_OF_DATE:INT
	VAR_INPUT
		IDATE :	UDINT;
	END_VAR

	YEAR_OF_DATE := UDINT_TO_INT((idate+UDINT#43200) / UDINT#31557600 + UDINT#1970);
END_FUNCTION

FUNCTION DT_TO_DATE2:UDINT

	VAR_INPUT
		IN :	UDINT;
	END_VAR

	DT_TO_DATE2 := (IN / UDINT#86400) * UDINT#86400;
END_FUNCTION

FUNCTION SET_DATE:UDINT

	VAR_INPUT
		YEAR :	INT;
		MONTH :	INT;
		DAY :	INT;
	END_VAR

	VAR
		count :	INT;
	END_VAR

	IF month > 2 THEN
		count := (month - 1) * 30;
		IF month > 7 THEN
			count := count + DWORD_TO_INT(SHR(DINT_TO_DWORD(INT_TO_DINT(month) - INT_TO_DINT(3)),1));
		ELSE
			count := count + DWORD_TO_INT(SHR(DINT_TO_DWORD(INT_TO_DINT(month) - INT_TO_DINT(4)),1));
		END_IF;
		IF SHL(INT_TO_WORD(year),14) = WORD#0 THEN
			count := count + 1;
		END_IF;
	ELSE
		count := (month - 1) * 31;
	END_IF;
	SET_DATE := (_INT_TO_UDINT(count + day - 1) + DWORD_TO_UDINT(SHR(UDINT_TO_DWORD(_INT_TO_UDINT(year) * UDINT#1461 - UDINT#2878169), 2))) * UDINT#86400;

END_FUNCTION

FUNCTION SET_DT:UDINT

	VAR_INPUT
		YEAR :	INT;
		MONTH :	INT;
		DAY :	INT;
		HOUR :	INT;
		MINUTE :	INT;
		SECOND :	INT;
	END_VAR

	SET_DT := SET_DATE(YEAR, MONTH, DAY) + _INT_TO_UDINT(SECOND) + _INT_TO_UDINT(MINUTE) * UDINT#60 + _INT_TO_UDINT(HOUR) * UDINT#3600;

END_FUNCTION

FUNCTION DST:BOOL
	VAR_INPUT
		UTC :	UDINT;
	END_VAR

	VAR
		yr :	INT;
		yr4 :	UDINT;
		ltc :	UDINT;
		idate :	UDINT;
	END_VAR

	yr := YEAR_OF_DATE(DT_TO_DATE2(UTC));
	ltc := UTC;
	idate := SET_DT(yr, 3, 31, 1, 0, 0);
	yr4 := DWORD_TO_UDINT(SHR(INT_TO_DWORD(5 * yr), 2)) + UDINT#1;
	DST := (idate - ((yr4 + UDINT#3) MOD UDINT#7) * UDINT#86400 <= ltc) AND (idate + (UDINT#214 - (yr4) MOD UDINT#7) * UDINT#86400 > ltc);
END_FUNCTION

PROGRAM program0
	VAR
		UTC :	UDINT;
		CEIL5_OUT : BOOL;
	END_VAR

  CEIL5_OUT := DST(UTC);

END_PROGRAM

CONFIGURATION Config0
	RESOURCE Res0 ON PLC
		TASK task0(INTERVAL := T#20ms,PRIORITY := 0);
		PROGRAM instance0 WITH task0 : program0;
	END_RESOURCE
END_CONFIGURATION

(* ---- DT_TO_DATE.ST ---- *)
FUNCTION _DT_TO_DATE_B:UDINT

	VAR_INPUT
		_INN :	UDINT;
	END_VAR

	_DT_TO_DATE_B := (_INN / UDINT#86400) * UDINT#86400;
END_FUNCTION

PROGRAM program0
	VAR
		_INN :	UDINT;
		OUT : UDINT;
	END_VAR

  OUT := _DT_TO_DATE_B(_INN);

CONFIGURATION Config0
	RESOURCE Res0 ON PLC
		TASK task0(INTERVAL := T#20ms,PRIORITY := 0);
		PROGRAM instance0 WITH task0 : program0;
	END_RESOURCE
END_CONFIGURATION

(* ---- DT_TO_TOD.ST ---- *)
FUNCTION DT_TO_TOD2:UDINT
	VAR_INPUT
		IN :	UDINT;
	END_VAR

	DT_TO_TOD2 := (IN MOD UDINT#86400) * UDINT#1000;
END_FUNCTION

PROGRAM program0
  VAR
    LocalVar0 : UDINT;
	LocalOUT  : UDINT;
  END_VAR
  	LocalOUT := DT_TO_TOD2(LocalVar0);
END_PROGRAM

CONFIGURATION Config0
  RESOURCE Res0 ON PLC
    TASK task0(INTERVAL := T#20ms,PRIORITY := 0);
    PROGRAM instance0 WITH task0 : program0;
  END_RESOURCE
END_CONFIGURATION

(* ---- DWORD_OF_BYTE.ST ---- *)
FUNCTION DWORD_OF_BYTE:DWORD
	VAR_INPUT
		B3 :	BYTE;
		B2 :	BYTE;
		B1 :	BYTE;
		B0 :	BYTE;
	END_VAR

	DWORD_OF_BYTE := SHL(SHL(SHL(BYTE_TO_DWORD(B3),8) OR BYTE_TO_DWORD(B2),8) OR BYTE_TO_DWORD(B1),8) OR BYTE_TO_DWORD(B0);

END_FUNCTION

PROGRAM program0
  VAR
    LocalVar0 : BYTE;
	LocalVar1 : BYTE;
	LocalVar2 : BYTE;
	LocalVar3 : BYTE;
	LocalOUT  : DWORD;
  END_VAR
  	LocalOUT := DWORD_OF_BYTE(LocalVar0, LocalVar1, LocalVar2, LocalVar3);
END_PROGRAM

CONFIGURATION Config0
  RESOURCE Res0 ON PLC
    TASK task0(INTERVAL := T#20ms,PRIORITY := 0);
    PROGRAM instance0 WITH task0 : program0;
  END_RESOURCE
END_CONFIGURATION

(* ---- DWORD_OF_WORD.ST ---- *)
FUNCTION DWORD_OF_WORD:DWORD

	VAR_INPUT
		W1 :	WORD;
		W0 :	WORD;
	END_VAR

	DWORD_OF_WORD := SHL(WORD_TO_DWORD(W1),16) OR WORD_TO_DWORD(W0);

END_FUNCTION

PROGRAM program0
  VAR
    LocalVar0 : WORD;
	LocalVar1 : WORD;
	LocalOUT  : DWORD;
  END_VAR
  	LocalOUT := DWORD_OF_WORD(LocalVar0, LocalVar1);
END_PROGRAM

CONFIGURATION Config0
  RESOURCE Res0 ON PLC
    TASK task0(INTERVAL := T#20ms,PRIORITY := 0);
    PROGRAM instance0 WITH task0 : program0;
  END_RESOURCE
END_CONFIGURATION

(* ---- DWORD_TO_DATE.ST ---- *)
FUNCTION DWORD_TO_DATE2:UDINT
	VAR_INPUT
		IN :	DWORD;
	END_VAR
	DWORD_TO_DATE2 := DWORD_TO_UDINT(IN);
END_FUNCTION

PROGRAM program0
  VAR
    LocalVar0 : DWORD;
	LocalOUT  : UDINT;
  END_VAR
  	LocalOUT := DWORD_TO_DATE2(LocalVar0);
END_PROGRAM

CONFIGURATION Config0
  RESOURCE Res0 ON PLC
    TASK task0(INTERVAL := T#20ms,PRIORITY := 0);
    PROGRAM instance0 WITH task0 : program0;
  END_RESOURCE
END_CONFIGURATION

(* ---- DWORD_TO_DT.ST ---- *)
FUNCTION DWORD_TO_DT2:UDINT

	VAR_INPUT
		IN :	DWORD;
	END_VAR

	DWORD_TO_DT2 := DWORD_TO_UDINT(IN);
END_FUNCTION

PROGRAM program0
  VAR
    LocalVar0 : DWORD;
	LocalOUT  : UDINT;
  END_VAR
  	LocalOUT := DWORD_TO_DT2(LocalVar0);
END_PROGRAM

CONFIGURATION Config0
  RESOURCE Res0 ON PLC
    TASK task0(INTERVAL := T#20ms,PRIORITY := 0);
    PROGRAM instance0 WITH task0 : program0;
  END_RESOURCE
END_CONFIGURATION

(* ---- DWORD_TO_TIME.ST ---- *)
FUNCTION DWORD_TO_TIME2:TIME
	VAR_INPUT
		X :	DWORD;
	END_VAR
	DWORD_TO_TIME2 := DINT_TO_TIME(DWORD_TO_DINT(X));
END_FUNCTION

PROGRAM program0
  VAR
    LocalVar0 : DWORD;
	  LocalOUT  : TIME;
  END_VAR
  	LocalOUT := DWORD_TO_TIME2(LocalVar0);
END_PROGRAM

CONFIGURATION Config0
  RESOURCE Res0 ON PLC
    TASK task0(INTERVAL := T#20ms,PRIORITY := 0);
    PROGRAM instance0 WITH task0 : program0;
  END_RESOURCE
END_CONFIGURATION

(* ---- DWORD_TO_TOD.ST ---- *)
FUNCTION DWORD_TO_TOD2:UDINT
	VAR_INPUT
		IN :	DWORD;
	END_VAR
	DWORD_TO_TOD2 := DWORD_TO_UDINT(IN);
END_FUNCTION

PROGRAM program0
  VAR
    LocalVar0 : DWORD;
	  LocalOUT  : UDINT;
  END_VAR
  	LocalOUT := DWORD_TO_TOD2(LocalVar0);
END_PROGRAM

CONFIGURATION Config0
  RESOURCE Res0 ON PLC
    TASK task0(INTERVAL := T#20ms,PRIORITY := 0);
    PROGRAM instance0 WITH task0 : program0;
  END_RESOURCE
END_CONFIGURATION

(* ---- EASTER.ST ---- *)
FUNCTION _INT_TO_UDINT:UDINT
	VAR_INPUT
		IN :	INT;
	END_VAR

	_INT_TO_UDINT := DINT_TO_UDINT(INT_TO_DINT(IN));
END_FUNCTION

FUNCTION SET_DATE:UDINT

	VAR_INPUT
		YEAR :	INT;
		MONTH :	INT;
		DAY :	INT;
	END_VAR

	VAR
		count :	INT;
	END_VAR

	IF month > 2 THEN
		count := (month - 1) * 30;
		IF month > 7 THEN
			count := count + DWORD_TO_INT(SHR(DINT_TO_DWORD(INT_TO_DINT(month) - INT_TO_DINT(3)),1));
		ELSE
			count := count + DWORD_TO_INT(SHR(DINT_TO_DWORD(INT_TO_DINT(month) - INT_TO_DINT(4)),1));
		END_IF;
		IF SHL(INT_TO_WORD(year),14) = WORD#0 THEN
			count := count + 1;
		END_IF;
	ELSE
		count := (month - 1) * 31;
	END_IF;
	SET_DATE := (_INT_TO_UDINT(count + day - 1) + DWORD_TO_UDINT(SHR(UDINT_TO_DWORD(_INT_TO_UDINT(year) * UDINT#1461 - UDINT#2878169), 2))) * UDINT#86400;

END_FUNCTION

FUNCTION EASTER:UDINT
	VAR_INPUT
		YEAR :	INT;
	END_VAR

	VAR
		b :	INT;
		c :	INT;
		oday :	INT;
	END_VAR

	b := (204 - 11 * (year MOD 19)) MOD 30;
	IF b > 27 THEN b := b - 1; END_IF;
	c := (year + WORD_TO_INT(SHR(INT_TO_WORD(year),2)) + b - 13) MOD 7;
	oday := 28 + b - c;
	IF oday > 33 THEN
		easter := set_Date(year, 4, oday - 31);
	ELSE
		easter := set_Date(year, 3, oday);
	END_IF;
END_FUNCTION

PROGRAM program0
  VAR
    LocalVar0 : INT;
	LocalOUT  : UDINT;
  END_VAR
  	LocalOUT := EASTER(LocalVar0);
END_PROGRAM

CONFIGURATION Config0
  RESOURCE Res0 ON PLC
    TASK task0(INTERVAL := T#20ms,PRIORITY := 0);
    PROGRAM instance0 WITH task0 : program0;
  END_RESOURCE
END_CONFIGURATION

(* ---- ELLIPSE_A.ST ---- *)
FUNCTION ELLIPSE_A:REAL
	VAR_INPUT
		R1 :	REAL;
		R2 :	REAL;
	END_VAR

	ellipse_A := 3.14159265358979323846264338327950288 * R1 * R2;

END_FUNCTION

PROGRAM program0
  VAR
    LocalVar0 : REAL;
	LocalVar1 : REAL;
	  LocalOUT  : REAL;
  END_VAR
  	LocalOUT := ELLIPSE_A(LocalVar0, LocalVar1);
END_PROGRAM

CONFIGURATION Config0
  RESOURCE Res0 ON PLC
    TASK task0(INTERVAL := T#20ms,PRIORITY := 0);
    PROGRAM instance0 WITH task0 : program0;
  END_RESOURCE
END_CONFIGURATION

(* ---- ELLIPSE_C.ST ---- *)
FUNCTION ELLIPSE_C:REAL

VAR_INPUT
	R1 :	REAL;
	R2 :	REAL;
END_VAR

ELLIPSE_C := 3.14159265358979323846264338327950288 * (3.0 * (R1+R2) - SQRT((3.0 * r1 + R2) * (3.0 * r2 + r1)));

END_FUNCTION

PROGRAM program0
  VAR
    LocalVar0 : REAL;
	LocalVar1 : REAL;
	  LocalOUT  : REAL;
  END_VAR
  	LocalOUT := ELLIPSE_C(LocalVar0, LocalVar1);
END_PROGRAM

CONFIGURATION Config0
  RESOURCE Res0 ON PLC
    TASK task0(INTERVAL := T#20ms,PRIORITY := 0);
    PROGRAM instance0 WITH task0 : program0;
  END_RESOURCE
END_CONFIGURATION

(* ---- ERF.ST ---- *)
FUNCTION SGN : INT
  VAR_INPUT
    x : REAL;
  END_VAR

  IF X > 0.0 THEN
  	sgn := 1;
  ELSIF X < 0.0 THEN
  	sgn := -1;
  ELSE
  	sgn := 0;
  END_IF;
END_FUNCTION

FUNCTION ERF:REAL

	VAR_INPUT
		X :	REAL;
	END_VAR

	VAR
		x2 :	REAL;
		ax2 :	REAL;
	END_VAR

	x2 := X*X;
	ax2 := 0.147 * x2 + 1.0;
	ERF := SQRT(1.0 - EXP(-X2 * ((0.27323954473516 + aX2)/(ax2)))) * INT_TO_REAL(SGN(x));

END_FUNCTION

PROGRAM program0
  VAR
    LocalVar0 : REAL;
	  LocalOUT  : REAL;
  END_VAR
  	LocalOUT := ERF(LocalVar0);
END_PROGRAM

CONFIGURATION Config0
  RESOURCE Res0 ON PLC
    TASK task0(INTERVAL := T#20ms,PRIORITY := 0);
    PROGRAM instance0 WITH task0 : program0;
  END_RESOURCE
END_CONFIGURATION

(* ---- ERFC.ST ---- *)
FUNCTION SGN : INT
  VAR_INPUT
    x : REAL;
  END_VAR

  IF X > 0.0 THEN
  	sgn := 1;
  ELSIF X < 0.0 THEN
  	sgn := -1;
  ELSE
  	sgn := 0;
  END_IF;
END_FUNCTION

FUNCTION ERF:REAL

	VAR_INPUT
		X :	REAL;
	END_VAR

	VAR
		x2 :	REAL;
		ax2 :	REAL;
	END_VAR

	x2 := X*X;
	ax2 := 0.147 * x2 + 1.0;
	ERF := SQRT(1.0 - EXP(-X2 * ((0.27323954473516 + aX2)/(ax2)))) * INT_TO_REAL(SGN(x));

END_FUNCTION

FUNCTION ERFC:REAL
	VAR_INPUT
		X :	REAL;
	END_VAR

	ERFC := 1.0 - ERF(X);

END_FUNCTION

PROGRAM program0
  VAR
    LocalVar0 : REAL;
	  LocalOUT  : REAL;
  END_VAR
  	LocalOUT := ERFC(LocalVar0);
END_PROGRAM

CONFIGURATION Config0
  RESOURCE Res0 ON PLC
    TASK task0(INTERVAL := T#20ms,PRIORITY := 0);
    PROGRAM instance0 WITH task0 : program0;
  END_RESOURCE
END_CONFIGURATION

(* ---- EVEN.ST ---- *)
FUNCTION BIT_OF_DWORD : BOOL
  VAR_INPUT
    IN : DWORD;
    N : INT;
  END_VAR

  BIT_OF_DWORD := (SHR(in,N) AND 16#00000001) > 0;
END_FUNCTION

FUNCTION EVEN:BOOL
	VAR_INPUT
		IN :	DINT;
	END_VAR

	even := NOT BIT_OF_DWORD(DINT_TO_DWORD(in),0);
END_FUNCTION

PROGRAM program0
  VAR
    LocalVar0 : DINT;
	  LocalOUT  : BOOL;
  END_VAR
  	LocalOUT := EVEN(LocalVar0);
END_PROGRAM

CONFIGURATION Config0
  RESOURCE Res0 ON PLC
    TASK task0(INTERVAL := T#20ms,PRIORITY := 0);
    PROGRAM instance0 WITH task0 : program0;
  END_RESOURCE
END_CONFIGURATION

(* ---- EXP10.ST ---- *)
FUNCTION EXP10 : REAL
  VAR_INPUT
    x : REAL;
  END_VAR

  exp10 := EXP(X * 2.30258509299405);
  (* from OSCAT library; www.oscat.de  *)
END_FUNCTION

PROGRAM program0
  VAR
    LocalVar0 : REAL;
    CEIL5_OUT : REAL;
  END_VAR

  CEIL5_OUT := EXP10(LocalVar0);
END_PROGRAM

CONFIGURATION Config0

  RESOURCE Res0 ON PLC
    TASK task0(INTERVAL := T#20ms,PRIORITY := 0);
    PROGRAM instance0 WITH task0 : program0;
  END_RESOURCE
END_CONFIGURATION

(* ---- EXPN.ST ---- *)
FUNCTION BIT_OF_DWORD : BOOL
  VAR_INPUT
    IN : DWORD;
    N : INT;
  END_VAR

  BIT_OF_DWORD := (SHR(in,N) AND 16#00000001) > 0;
END_FUNCTION

FUNCTION EXPN:REAL

	VAR_INPUT
		X :	REAL;
		N :	INT;
	END_VAR

	VAR
		N_word :	WORD;
		X_tmp :	REAL;
		sign :	BOOL;
	END_VAR

	N_word := INT_TO_WORD(N);
	X_tmp := X;
	sign := BIT_OF_DWORD(WORD_TO_DWORD(N_word),15);
	N_word := INT_TO_WORD(ABS(N));
	IF BIT_OF_DWORD(WORD_TO_DWORD(N_word),0) THEN expn := X_tmp; ELSE expn := 1.0; END_IF;    (* N_word.X0 *)
	N_word := SHR(N_word,1);
	WHILE N_word > WORD#0 DO
		X_tmp := X_tmp * X_tmp;
		IF BIT_OF_DWORD(WORD_TO_DWORD(N_word),0) THEN expn := expn * X_tmp; END_IF;       (* N_word.X0 *)
		N_word := SHR(N_word,1);
	END_WHILE;
	IF sign THEN EXPN := 1.0 / EXPN; END_IF;

END_FUNCTION

PROGRAM program0
  VAR
    LocalVar0 : REAL;
	LocalVar1 : INT;
	LocalOUT  : REAL;
  END_VAR
  	LocalOUT := EXPN(LocalVar0, LocalVar1);
END_PROGRAM

CONFIGURATION Config0
  RESOURCE Res0 ON PLC
    TASK task0(INTERVAL := T#20ms,PRIORITY := 0);
    PROGRAM instance0 WITH task0 : program0;
  END_RESOURCE
END_CONFIGURATION

(* ---- F_LIN.ST ---- *)
FUNCTION F_LIN:REAL
	VAR_INPUT
		X :	REAL;
		A :	REAL;
		B :	REAL;
	END_VAR

	F_lin := A * X + B;
END_FUNCTION

PROGRAM program0
  VAR
    LocalVar0 : REAL;
	LocalVar1 : REAL;
	LocalVar2 : REAL;
	  LocalOUT  : REAL;
  END_VAR
  	LocalOUT := F_LIN(LocalVar0, LocalVar1, LocalVar2);
END_PROGRAM

CONFIGURATION Config0
  RESOURCE Res0 ON PLC
    TASK task0(INTERVAL := T#20ms,PRIORITY := 0);
    PROGRAM instance0 WITH task0 : program0;
  END_RESOURCE
END_CONFIGURATION

(* ---- F_LIN2.ST ---- *)
FUNCTION F_LIN2:REAL
	VAR_INPUT
		X :	REAL;
		X1 :	REAL;
		Y1 :	REAL;
		X2 :	REAL;
		Y2 :	REAL;
	END_VAR

	F_LIN2 := (Y2 - Y1) / (X2 - X1) * (X - X1) + Y1;

END_FUNCTION

PROGRAM program0
  VAR
    LocalVar0 : REAL;
	LocalVar1 : REAL;
	LocalVar2 : REAL;
	LocalVar3 : REAL;
	LocalVar4 : REAL;
	  LocalOUT  : REAL;
  END_VAR
  	LocalOUT := F_LIN2(LocalVar0, LocalVar1, LocalVar2, LocalVar3, LocalVar4);
END_PROGRAM

CONFIGURATION Config0
  RESOURCE Res0 ON PLC
    TASK task0(INTERVAL := T#20ms,PRIORITY := 0);
    PROGRAM instance0 WITH task0 : program0;
  END_RESOURCE
END_CONFIGURATION

(* ---- F_POWER.ST ---- *)
FUNCTION F_POWER:REAL
	VAR_INPUT
		A :	REAL;
		X :	REAL;
		N :	REAL;
	END_VAR

	f_power := a * EXPT(X,N);
END_FUNCTION

PROGRAM program0
  VAR
    LocalVar0 : REAL;
	LocalVar1 : REAL;
	LocalVar2 : REAL;
	  LocalOUT  : REAL;
  END_VAR
  	LocalOUT := F_POWER(LocalVar0, LocalVar1, LocalVar2);
END_PROGRAM

CONFIGURATION Config0
  RESOURCE Res0 ON PLC
    TASK task0(INTERVAL := T#20ms,PRIORITY := 0);
    PROGRAM instance0 WITH task0 : program0;
  END_RESOURCE
END_CONFIGURATION

(* ---- F_QUAD.ST ---- *)
FUNCTION F_QUAD:REAL

	VAR_INPUT
		X :	REAL;
		A :	REAL;
		B :	REAL;
		C :	REAL;
	END_VAR

	F_QUAD :=  (A * X + B) * X + C;

END_FUNCTION

PROGRAM program0
  VAR
    LocalVar0 : REAL;
	LocalVar1 : REAL;
	LocalVar2 : REAL;
	LocalVar3 : REAL;
	LocalOUT  : REAL;
  END_VAR
  	LocalOUT := F_QUAD(LocalVar0, LocalVar1, LocalVar2, LocalVar3);
END_PROGRAM

CONFIGURATION Config0
  RESOURCE Res0 ON PLC
    TASK task0(INTERVAL := T#20ms,PRIORITY := 0);
    PROGRAM instance0 WITH task0 : program0;
  END_RESOURCE
END_CONFIGURATION

(* ---- F_TO_C.ST ---- *)
FUNCTION F_TO_C:REAL
	VAR_INPUT
		FAHRENHEIT :	REAL;
	END_VAR
	F_TO_C := (fahrenheit - 32.0) * 0.5555555555555;
END_FUNCTION

PROGRAM program0
  VAR
    LocalVar0 : REAL;
	LocalOUT  : REAL;
  END_VAR
  	LocalOUT := F_TO_C(LocalVar0);
END_PROGRAM

CONFIGURATION Config0
  RESOURCE Res0 ON PLC
    TASK task0(INTERVAL := T#20ms,PRIORITY := 0);
    PROGRAM instance0 WITH task0 : program0;
  END_RESOURCE
END_CONFIGURATION

(* ---- F_TO_OM.ST ---- *)
FUNCTION F_TO_OM:REAL

	VAR_INPUT
		F :	REAL;
	END_VAR

	F_to_OM := 6.283185307179586476 * F;

END_FUNCTION

PROGRAM program0
  VAR
    LocalVar0 : REAL;
	  LocalOUT  : REAL;
  END_VAR
  	LocalOUT := F_TO_OM(LocalVar0);
END_PROGRAM

CONFIGURATION Config0
  RESOURCE Res0 ON PLC
    TASK task0(INTERVAL := T#20ms,PRIORITY := 0);
    PROGRAM instance0 WITH task0 : program0;
  END_RESOURCE
END_CONFIGURATION

(* ---- F_TO_PT.ST ---- *)
FUNCTION _REAL_TO_DWORD: DWORD
  VAR_INPUT
    X :	REAL;
  END_VAR

  IF REAL_TO_DWORD(0.5) = DWORD#1 THEN
    _REAL_TO_DWORD := REAL_TO_DWORD(x);
  ELSIF X > 0.0 THEN
    _REAL_TO_DWORD := REAL_TO_DWORD(x+0.5);
  ELSIF X < 0.0 THEN
    _REAL_TO_DWORD := REAL_TO_DWORD(x-0.5);
  ELSE
    _REAL_TO_DWORD := DWORD#0;
  END_IF;
END_FUNCTION

FUNCTION F_TO_PT:TIME
	VAR_INPUT
		F :	REAL;
	END_VAR
	F_TO_PT := DWORD_TO_TIME(_REAL_TO_DWORD(1.0 / F * 1000.0));
END_FUNCTION

PROGRAM program0
  VAR
    LocalVar0 : REAL;
	  LocalOUT  : TIME;
  END_VAR
  	LocalOUT := F_TO_PT(LocalVar0);
END_PROGRAM

CONFIGURATION Config0
  RESOURCE Res0 ON PLC
    TASK task0(INTERVAL := T#20ms,PRIORITY := 0);
    PROGRAM instance0 WITH task0 : program0;
  END_RESOURCE
END_CONFIGURATION

(* ---- FACT.ST ---- *)
FUNCTION FACT:DINT

	VAR_INPUT
		X :	INT;
	END_VAR

	CASE X OF
	00: FACT := DINT#1;
	01: FACT := DINT#1;
	02: FACT := DINT#2;
	03: FACT := DINT#6;
	04: FACT := DINT#24;
	05: FACT := DINT#120;
	06: FACT := DINT#720;
	07: FACT := DINT#5040;
	08: FACT := DINT#40320;
	09: FACT := DINT#362880;
	10: FACT := DINT#3628800;
	11: FACT := DINT#39916800;
	12: FACT := DINT#479001600;
	ELSE
		FACT := DINT#-1;
	END_CASE;

END_FUNCTION

PROGRAM program0
  VAR
    LocalVar0 : INT;
	LocalOUT  : DINT;
  END_VAR
  	LocalOUT := FACT(LocalVar0);
END_PROGRAM

CONFIGURATION Config0
  RESOURCE Res0 ON PLC
    TASK task0(INTERVAL := T#20ms,PRIORITY := 0);
    PROGRAM instance0 WITH task0 : program0;
  END_RESOURCE
END_CONFIGURATION

(* ---- FIB.ST ---- *)
FUNCTION FIB:DINT

VAR_INPUT
	X :	INT;
END_VAR

VAR
	t1 :	DINT;
	t2 :	DINT;
	X_tmp :	INT;
END_VAR

t1 := DINT#0;
t2 := DINT#0;
X_tmp := X;
IF X_tmp < 0 OR X_tmp > 46 THEN
	FIB := DINT#-1;
ELSIF X_tmp < 2 THEN
	FIB := INT_TO_DINT(X_tmp);
	RETURN;
ELSE
	t2 := DINT#1;
	WHILE X_tmp > 3 DO
		X_tmp := X_tmp - 2;
		t1 := t1 + t2;
		t2 := t1 + t2;
	END_WHILE;
	IF X_tmp > 2 THEN t1 := t1 + t2; END_IF;
	fib := t1 + t2;
END_IF;

END_FUNCTION

PROGRAM program0
  VAR
    LocalVar0 : INT;
	LocalOUT  : DINT;
  END_VAR
  	LocalOUT := FIB(LocalVar0);
END_PROGRAM

CONFIGURATION Config0
  RESOURCE Res0 ON PLC
    TASK task0(INTERVAL := T#20ms,PRIORITY := 0);
    PROGRAM instance0 WITH task0 : program0;
  END_RESOURCE
END_CONFIGURATION

(* ---- FLOOR.ST ---- *)
FUNCTION FLOOR : INT
  VAR_INPUT
    x : REAL;
  END_VAR

  FLOOR := REAL_TO_INT(X);
  IF INT_TO_REAL(FLOOR) > X THEN
  	floor := floor - 1;
  END_IF;
  (* from OSCAT library; www.oscat.de  *)
END_FUNCTION

PROGRAM program0
  VAR
    LocalVar0 : REAL;
    CEIL5_OUT : INT;
  END_VAR

  CEIL5_OUT := FLOOR(LocalVar0);
END_PROGRAM

CONFIGURATION Config0

  RESOURCE Res0 ON PLC
    TASK task0(INTERVAL := T#20ms,PRIORITY := 0);
    PROGRAM instance0 WITH task0 : program0;
  END_RESOURCE
END_CONFIGURATION

(* ---- FLOOR2.ST ---- *)
FUNCTION _REAL_TO_DINT:DINT
  VAR_INPUT
    X :	REAL;
  END_VAR

  IF REAL_TO_DINT(0.5) = DINT#1 THEN
    _REAL_TO_DINT := REAL_TO_DINT(x);
    RETURN;
  END_IF;

  IF X > 0.0 THEN
    _REAL_TO_DINT := REAL_TO_DINT(x+0.5);
  ELSIF X < 0.0 THEN
    _REAL_TO_DINT := REAL_TO_DINT(x-0.5);
  ELSE
    _REAL_TO_DINT := DINT#0;
  END_IF;
END_FUNCTION

FUNCTION FLOOR2:DINT
	VAR_INPUT
		X :	REAL;
	END_VAR

	FLOOR2 := _REAL_TO_DINT(X);
	IF DINT_TO_REAL(FLOOR2) > X THEN
		FLOOR2 := FLOOR2 - DINT#1;
	END_IF;
END_FUNCTION

PROGRAM program0
  VAR
    LocalVar0 : REAL;
    CEIL5_OUT : DINT;
  END_VAR

  CEIL5_OUT := FLOOR2(LocalVar0);
END_PROGRAM

CONFIGURATION Config0

  RESOURCE Res0 ON PLC
    TASK task0(INTERVAL := T#20ms,PRIORITY := 0);
    PROGRAM instance0 WITH task0 : program0;
  END_RESOURCE
END_CONFIGURATION

(* ---- FRACT.ST ---- *)
FUNCTION D_TRUNC : DINT
  VAR_INPUT
    x : REAL;
  END_VAR

  D_TRUNC := REAL_TO_DINT(X);
  IF X > 0.0 THEN
  	IF DINT_TO_REAL(D_TRUNC) > X THEN D_TRUNC := D_TRUNC - DINT#1; END_IF;
  ELSE
  	IF DINT_TO_REAL(D_TRUNC) < X THEN D_TRUNC := D_TRUNC + DINT#1; END_IF;
  END_IF;
END_FUNCTION

FUNCTION FRACT:REAL
	VAR_INPUT
		X :	REAL;
	END_VAR

	IF ABS(x) < 2.0E9 THEN
		FRACT := x - DINT_TO_REAL(D_TRUNC(x));
	ELSE
		FRACT := 0.0;
	END_IF;
END_FUNCTION

PROGRAM program0
  VAR
    LocalVar0 : REAL;
	LocalOUT  : REAL;
  END_VAR
  	LocalOUT := FRACT(LocalVar0);
END_PROGRAM

CONFIGURATION Config0
  RESOURCE Res0 ON PLC
    TASK task0(INTERVAL := T#20ms,PRIORITY := 0);
    PROGRAM instance0 WITH task0 : program0;
  END_RESOURCE
END_CONFIGURATION

(* ---- FRMP_B.ST ---- *)
FUNCTION FRMP_B:BYTE

	VAR_INPUT
		START :	BYTE;
		DIR :	BOOL;
		TD :	TIME;
		TR :	TIME;
	END_VAR

	IF TD < TR THEN
		FRMP_B := MIN(UDINT_TO_BYTE(DWORD_TO_UDINT(SHL(TIME_TO_DWORD(TD), 8)) / TIME_TO_UDINT(TR)), SEL(DIR, START, USINT_TO_BYTE(USINT#255 - BYTE_TO_USINT(START))));
		IF DIR THEN
			FRMP_B := USINT_TO_BYTE(BYTE_TO_USINT(START) + BYTE_TO_USINT(FRMP_B));
		ELSE
			FRMP_B := USINT_TO_BYTE(BYTE_TO_USINT(START) - BYTE_TO_USINT(FRMP_B));
		END_IF;
	ELSE
		FRMP_B := SEL(DIR, BYTE#0, BYTE#255);
	END_IF;
END_FUNCTION

PROGRAM program0
  VAR
    LocalVar0 : BYTE;
	LocalVar1 : BOOL;
	LocalVar2 : TIME;
	LocalVar3 : TIME;
    LocalOUT  : BYTE;
  END_VAR

  LocalOUT := FRMP_B(LocalVar0, LocalVar1, LocalVar2,LocalVar3);
END_PROGRAM

CONFIGURATION Config0
  RESOURCE Res0 ON PLC
    TASK task0(INTERVAL := T#20ms,PRIORITY := 0);
    PROGRAM instance0 WITH task0 : program0;
  END_RESOURCE
END_CONFIGURATION

(* ---- GAMMA.ST ---- *)
FUNCTION GAMMA:REAL
	VAR_INPUT
		X :	REAL;
	END_VAR

	IF x > 0.0 THEN
		GAMMA := SQRT(6.28318530717958647692528676655900576 / X) * EXPT(0.367879441171442 * (x + 1.0 / (12.0 * x - 0.1 / X)), X);
	END_IF;
END_FUNCTION

PROGRAM program0
  VAR
    LocalVar0 : REAL;
    LocalOUT  : REAL;
  END_VAR

  LocalOUT := GAMMA(LocalVar0);
END_PROGRAM

CONFIGURATION Config0
  RESOURCE Res0 ON PLC
    TASK task0(INTERVAL := T#20ms,PRIORITY := 0);
    PROGRAM instance0 WITH task0 : program0;
  END_RESOURCE
END_CONFIGURATION

(* ---- GAUSS.ST ---- *)
FUNCTION GAUSS:REAL

	VAR_INPUT
		X :	REAL;
		U :	REAL;
		SI :	REAL;
	END_VAR

	VAR
		temp :	REAL;
		si_inv :	REAL;
	END_VAR

	temp := X - U;
	si_inv := 1.0  / si;
	GAUSS := EXP(Temp * Temp * si_inv * SI_inv * - 0.5) * 0.39894228 * si_inv;

END_FUNCTION

PROGRAM program0
  VAR
    X :	REAL;
	U :	REAL;
	SI :	REAL;
    LocalOUT  : REAL;
  END_VAR

  LocalOUT := GAUSS(X, U, SI);
END_PROGRAM

CONFIGURATION Config0
  RESOURCE Res0 ON PLC
    TASK task0(INTERVAL := T#20ms,PRIORITY := 0);
    PROGRAM instance0 WITH task0 : program0;
  END_RESOURCE
END_CONFIGURATION

(* ---- GAUSSCD.ST ---- *)
FUNCTION SGN : INT
  VAR_INPUT
    x : REAL;
  END_VAR

  IF X > 0.0 THEN
  	sgn := 1;
  ELSIF X < 0.0 THEN
  	sgn := -1;
  ELSE
  	sgn := 0;
  END_IF;
END_FUNCTION

FUNCTION ERF:REAL

	VAR_INPUT
		X :	REAL;
	END_VAR

	VAR
		x2 :	REAL;
		ax2 :	REAL;
	END_VAR

	x2 := X*X;
	ax2 := 0.147 * x2 + 1.0;
	ERF := SQRT(1.0 - EXP(-X2 * ((0.27323954473516 + aX2)/(ax2)))) * INT_TO_REAL(SGN(x));

END_FUNCTION

FUNCTION GAUSSCD:REAL

	VAR_INPUT
		X :	REAL;
		U :	REAL;
		SI :	REAL;
	END_VAR

	GAUSSCD := (ERF((X - U) / (SI * 1.414213562)) + 1.0) * 0.5;

END_FUNCTION

PROGRAM program0
  VAR
    X :	REAL;
	U :	REAL;
	SI :	REAL;
    LocalOUT  : REAL;
  END_VAR

  LocalOUT := GAUSSCD(X, U, SI);
END_PROGRAM

CONFIGURATION Config0
  RESOURCE Res0 ON PLC
    TASK task0(INTERVAL := T#20ms,PRIORITY := 0);
    PROGRAM instance0 WITH task0 : program0;
  END_RESOURCE
END_CONFIGURATION

(* ---- GCD.ST ---- *)
FUNCTION GCD:INT

	VAR_INPUT
		A :	DINT;
		B :	DINT;
	END_VAR

	VAR
		t :	DINT;
		_A :	DINT;
		_B :	DINT;
	END_VAR

	_A := A;
	_B := B;

	IF _A = DINT#0 THEN
		GCD := DINT_TO_INT(ABS(_B));
	ELSIF _B = DINT#0 THEN
		GCD := DINT_TO_INT(ABS(_A));
	ELSE
		_A := ABS(_A);
		_B := ABS(_B);
		GCD := 1;

		WHILE NOT((DINT_TO_DWORD(_A) AND DWORD#1) > DWORD#0 OR (DINT_TO_DWORD(_B) AND DWORD#1) > DWORD#0) DO
			_A := DWORD_TO_DINT(SHR(DINT_TO_DWORD(_A),1));
			_B := DWORD_TO_DINT(SHR(DINT_TO_DWORD(_B),1));
			GCD := DWORD_TO_INT(SHR(INT_TO_DWORD(GCD),1));
		END_WHILE;
		WHILE _A > DINT#0 DO
			IF NOT((DINT_TO_DWORD(_A) AND DWORD#1) > DWORD#0) THEN
				_A := DWORD_TO_DINT(SHR(DINT_TO_DWORD(_A),1));
			ELSIF NOT((DINT_TO_DWORD(_B) AND DWORD#1) > DWORD#0) THEN
				_B := DWORD_TO_DINT(SHR(DINT_TO_DWORD(_B),1));
			ELSE
				t := DWORD_TO_DINT(SHR(DINT_TO_DWORD(ABS(_A-_B)),1));
				IF _A < _B THEN
					_B := t;
				ELSE
					_A := t;
				END_IF;
			END_IF;
		END_WHILE;
		GCD := GCD * DINT_TO_INT(_B);
	END_IF;

END_FUNCTION

PROGRAM program0
  VAR
    A :	DINT;
	B :	DINT;
    LocalOUT  : INT;
  END_VAR

  LocalOUT := GCD(A, B);
END_PROGRAM

CONFIGURATION Config0
  RESOURCE Res0 ON PLC
    TASK task0(INTERVAL := T#20ms,PRIORITY := 0);
    PROGRAM instance0 WITH task0 : program0;
  END_RESOURCE
END_CONFIGURATION

(* ---- GDF.ST ---- *)
FUNCTION GDF:REAL

	VAR_INPUT
		X :	REAL;
	END_VAR

	IF X = 0.0 THEN
		GDF := 0.0;
	ELSIF X > 15.0 THEN
		GDF := 1.5707963267949;
	ELSIF X < -15.0 THEN
		GDF := -1.5707963267949;
	ELSE
		GDF := ATAN(EXP(X)) * 2.0 - 1.5707963267949;
	END_IF;

END_FUNCTION

PROGRAM program0
  VAR
    X :	REAL;
    LocalOUT  : REAL;
  END_VAR

  LocalOUT := GDF(X);
END_PROGRAM

CONFIGURATION Config0
  RESOURCE Res0 ON PLC
    TASK task0(INTERVAL := T#20ms,PRIORITY := 0);
    PROGRAM instance0 WITH task0 : program0;
  END_RESOURCE
END_CONFIGURATION

(* ---- GEO_TO_DEG.ST ---- *)
FUNCTION GEO_TO_DEG:REAL

	VAR_INPUT
		D :	INT;
		M :	INT;
		SEC :	REAL;
	END_VAR

	GEO_TO_DEG := INT_TO_REAL(D) + INT_TO_REAL(M) * 0.016666666666667 + sec * 0.00027777777777778;

END_FUNCTION

PROGRAM program0
  VAR
    D :	INT;
	M :	INT;
	SEC :	REAL;
    LocalOUT  : REAL;
  END_VAR

  LocalOUT := GEO_TO_DEG(D, M, SEC);
END_PROGRAM

CONFIGURATION Config0
  RESOURCE Res0 ON PLC
    TASK task0(INTERVAL := T#20ms,PRIORITY := 0);
    PROGRAM instance0 WITH task0 : program0;
  END_RESOURCE
END_CONFIGURATION

(* ---- GOLD.ST ---- *)
FUNCTION GOLD:REAL

	VAR_INPUT
		X :	REAL;
	END_VAR

	GOLD := (X + SQRT(X*X + 4.0)) * 0.5;

END_FUNCTION

PROGRAM program0
  VAR
   	X :	REAL;
    LocalOUT  : REAL;
  END_VAR

  LocalOUT := GOLD(X);
END_PROGRAM

CONFIGURATION Config0
  RESOURCE Res0 ON PLC
    TASK task0(INTERVAL := T#20ms,PRIORITY := 0);
    PROGRAM instance0 WITH task0 : program0;
  END_RESOURCE
END_CONFIGURATION

(* ---- GRAY_TO_BYTE.ST ---- *)
FUNCTION GRAY_TO_BYTE:BYTE

	VAR_INPUT
		IN :	BYTE;
	END_VAR

	GRAY_TO_BYTE := SHR(IN,4) XOR IN;
	GRAY_TO_BYTE := SHR(GRAY_TO_BYTE,2) XOR GRAY_TO_BYTE;
	GRAY_TO_BYTE := SHR(GRAY_TO_BYTE,1) XOR GRAY_TO_BYTE;

END_FUNCTION

PROGRAM program0
  VAR
   	IN :	BYTE;
    LocalOUT  : BYTE;
  END_VAR

  LocalOUT := GRAY_TO_BYTE(IN);
END_PROGRAM

CONFIGURATION Config0
  RESOURCE Res0 ON PLC
    TASK task0(INTERVAL := T#20ms,PRIORITY := 0);
    PROGRAM instance0 WITH task0 : program0;
  END_RESOURCE
END_CONFIGURATION

(* ---- HEAT_INDEX.ST ---- *)
FUNCTION C_TO_F:REAL
	VAR_INPUT
		CELSIUS :	REAL;
	END_VAR

	C_TO_F := celsius * 1.8 + 32.0;
END_FUNCTION

FUNCTION F_TO_C:REAL
	VAR_INPUT
		FAHRENHEIT :	REAL;
	END_VAR
	F_TO_C := (fahrenheit - 32.0) * 0.5555555555555;
END_FUNCTION

FUNCTION HEAT_INDEX:REAL

	VAR_INPUT
		T :	REAL;
		RH :	REAL;
	END_VAR

	VAR
		RH2 :	REAL;
		T2 :	REAL;
		TX :	REAL;
	END_VAR

	IF RH < 20.0 OR T < 20.0 THEN
		HEAT_INDEX := T;
	ELSE
		TX := T;
		RH2 := RH * RH;
		TX := C_TO_F(TX);
		T2 := TX * TX;
		HEAT_INDEX := -42.379 + 2.04901523 * TX - 6.83783E-3 * T2
				+ RH * (10.1433127 - 0.22475541 * TX + 1.22874E-3 * T2)
				+ RH2 * (8.5282E-4 * TX - 5.481717E-2 - 1.99E-6 * T2);
		HEAT_INDEX := F_TO_C(HEAT_INDEX);
	END_IF;

END_FUNCTION

PROGRAM program0
  VAR
    T :	REAL;
	RH :	REAL;
    CEIL5_OUT : REAL;
  END_VAR

  CEIL5_OUT := HEAT_INDEX(T, RH);
END_PROGRAM

CONFIGURATION Config0

  RESOURCE Res0 ON PLC
    TASK task0(INTERVAL := T#20ms,PRIORITY := 0);
    PROGRAM instance0 WITH task0 : program0;
  END_RESOURCE
END_CONFIGURATION

(* ---- HOUR.ST ---- *)
FUNCTION HOUR:INT
	VAR_INPUT
		ITOD :	UDINT;
	END_VAR
	hour := UDINT_TO_INT(itod / UDINT#3600000);
END_FUNCTION

PROGRAM program0
  VAR
	  ITOD :	UDINT;
    CEIL5_OUT : INT;
  END_VAR

  CEIL5_OUT := HOUR(ITOD);
END_PROGRAM

CONFIGURATION Config0

  RESOURCE Res0 ON PLC
    TASK task0(INTERVAL := T#20ms,PRIORITY := 0);
    PROGRAM instance0 WITH task0 : program0;
  END_RESOURCE
END_CONFIGURATION

(* ---- HOUR_OF_DT.ST ---- *)
FUNCTION HOUR_OF_DT:INT
	VAR_INPUT
		XDT :	UDINT;
	END_VAR

	HOUR_OF_DT := UDINT_TO_INT((XDT MOD UDINT#86400) / UDINT#3600);
END_FUNCTION

PROGRAM program0
  VAR
    LocalVar0 : UDINT;
	LocalOUT  : INT;
  END_VAR
  	LocalOUT := HOUR_OF_DT(LocalVar0);
END_PROGRAM

CONFIGURATION Config0
  RESOURCE Res0 ON PLC
    TASK task0(INTERVAL := T#20ms,PRIORITY := 0);
    PROGRAM instance0 WITH task0 : program0;
  END_RESOURCE
END_CONFIGURATION

(* ---- HOUR_TO_TIME.ST ---- *)
FUNCTION _REAL_TO_UDINT:UDINT
	VAR_INPUT
		X :	REAL;
	END_VAR

	IF REAL_TO_UDINT(0.5) = UDINT#1 THEN
		_REAL_TO_UDINT := REAL_TO_UDINT(x);
	ELSIF X > 0.0 THEN
		_REAL_TO_UDINT := REAL_TO_UDINT(x+0.5);
	ELSIF X < 0.0 THEN
		_REAL_TO_UDINT := REAL_TO_UDINT(x-0.5);
	ELSE
		_REAL_TO_UDINT := UDINT#0;
  	END_IF;
END_FUNCTION

FUNCTION HOUR_TO_TIME:TIME

	VAR_INPUT
		IN :	REAL;
	END_VAR

	hour_to_time := UDINT_TO_TIME(_REAL_TO_UDINT(IN * 3600000.0));

END_FUNCTION

PROGRAM program0

	VAR
		IN :	REAL;
		CEIL5_OUT : TIME;
	END_VAR

  	CEIL5_OUT := HOUR_TO_TIME(IN);

END_PROGRAM

CONFIGURATION Config0

	RESOURCE Res0 ON PLC
		TASK task0(INTERVAL := T#20ms,PRIORITY := 0);
		PROGRAM instance0 WITH task0 : program0;
	END_RESOURCE

END_CONFIGURATION

(* ---- HOUR_TO_TOD.ST ---- *)
FUNCTION _REAL_TO_UDINT:UDINT
	VAR_INPUT
		X :	REAL;
	END_VAR

	IF REAL_TO_UDINT(0.5) = UDINT#1 THEN
		_REAL_TO_UDINT := REAL_TO_UDINT(x);
	ELSIF X > 0.0 THEN
		_REAL_TO_UDINT := REAL_TO_UDINT(x+0.5);
	ELSIF X < 0.0 THEN
		_REAL_TO_UDINT := REAL_TO_UDINT(x-0.5);
	ELSE
		_REAL_TO_UDINT := UDINT#0;
	END_IF;

END_FUNCTION

FUNCTION HOUR_TO_TOD:UDINT

	VAR_INPUT
		IN :	REAL;
	END_VAR

	hour_to_tod := _REAL_TO_UDINT(IN * 3600000.00);

END_FUNCTION

PROGRAM program0
	VAR
		IN :	REAL;
		CEIL5_OUT : UDINT;
	END_VAR

  	CEIL5_OUT := HOUR_TO_TOD(IN);
END_PROGRAM

CONFIGURATION Config0

  RESOURCE Res0 ON PLC
    TASK task0(INTERVAL := T#20ms,PRIORITY := 0);
    PROGRAM instance0 WITH task0 : program0;
  END_RESOURCE

END_CONFIGURATION

(* ---- HYPOT.ST ---- *)
FUNCTION HYPOT:REAL
	VAR_INPUT
		X :	REAL;
		Y :	REAL;
	END_VAR

	HYPOT := SQRT(x*x + y*y);
END_FUNCTION

PROGRAM program0
  VAR
    LocalVar0 : REAL;
    LocalVar1 : REAL;
    CEIL5_OUT : REAL;
  END_VAR

  CEIL5_OUT := HYPOT(LocalVar0, LocalVar1);
END_PROGRAM

CONFIGURATION Config0

  RESOURCE Res0 ON PLC
    TASK task0(INTERVAL := T#20ms,PRIORITY := 0);
    PROGRAM instance0 WITH task0 : program0;
  END_RESOURCE
END_CONFIGURATION
